// TIA Portal project "2023546359" (V18)

(* hardware
DEVICE "S7-1200 station_1"  S7-1200 Station
   slot 0: "Rack_0"  S7-1200 Rack  Rack  V1.0
   slot 1: "PLC"  CPU 1214C DC/DC/DC  6ES7 214-1AG40-0XB0  V4.2
*)

// ===== PLC "PLC"  CPU 1214C DC/DC/DC =====

VAR_GLOBAL CONSTANT   // PLC tag table "常量表"
   "ELE_SUM" : Int := 6;   // 电梯数量
   "FlOOR_TOP" : Int := 10;   // 电梯楼层
   "STATIC" : Int := 0;   // 静止状态
   "UP_H" : Int := 1;   // 上行高速
   "UP_L" : Int := 2;   // 上行低速
   "DOWN_H" : Int := 3;   // 下行高速
   "DOWN_L" : Int := 4;   // 下行低速
   "OPEN" : Int := 5;   // 开门
   "CLOSE" : Int := 6;   // 关门
   "H_L" : Int := 7;   // 高速转低速
   "L_H" : Int := 8;   // 低速转高速
   "SET_ELE" : Int := 5;
   "SET_FLOOR" : Int := 8;
END_VAR

TYPE "Button_Group"
   STRUCT
      state : Bool;
      light : Bool;
      p : Bool;
   END_STRUCT;
END_TYPE

TYPE "Elevator_Group"
   STRUCT
      jinggao : Struct
         REP : Bool;
         LC : Bool;
      END_STRUCT;
      display : Struct
         light : Bool;
         fan : Bool;
         error : Bool;
         full : Bool;
      END_STRUCT;
      direction : Struct
         up : Bool;
         down : Bool;
      END_STRUCT;
      door_jdq : Struct
         open : Bool;
         close : Bool;
      END_STRUCT;
      door_inplace : Struct
         close : Bool;
         open : Bool;
      END_STRUCT;
      bt_limit : Struct
         top1 : Bool;
         top2 : Bool;
         bottom1 : Bool;
         bottom2 : Bool;
      END_STRUCT;
      smg : Array[1..2, 1..7] of Bool;
      ele_speed : Struct
         H : Bool;
         L : Bool;
      END_STRUCT;
      run_contactor : Struct
         up : Bool;
         dowm : Bool;
      END_STRUCT;
      run_disp : Struct
         up : Bool;
         dowm : Bool;
      END_STRUCT;
      Brake : Struct
         B1 : Bool;
         B2 : Bool;
         B3 : Bool;
      END_STRUCT;
      floor_Lock : Array[1.."FlOOR_TOP"] of Bool;
      door_Lock : Bool;
      door_open : "Button_Group";
      btn_close : "Button_Group";
      ele_in_button : Array[1.."FlOOR_TOP"] of "Button_Group";
      run_enable : Bool;
      zhongliang : Word;
      button_out : Array[1..2, 1.."FlOOR_TOP"] of "Button_Group";   // 公共外部按键
   END_STRUCT;
END_TYPE

TYPE "Variable_Group"
   STRUCT
      init : Struct   // 初始化相关变量
         Init_state : Int;   // 初始化状态机
         kaishi : Bool;   // 初始化开始信号
         Init_now_f : Int;   // 初始化当前楼层
         mubiao_floor : Int;   // 初始化目标楼层
         init_fangxiang : Bool;   // 初始化方向
         jieshu : Bool;
         re_fangxiang : Bool;   // 检修后初始化方向
         re_mode : Bool;   // 检修后初始化方向设置模式(0自动1手动)
      END_STRUCT;
      Floor_handle : Struct   // 楼层处理相关变量
         dangqian_floor : Int;   // 当前楼层
         tag_1 : Bool;
         tag_2 : Bool;
      END_STRUCT;
      Weight_handle : Struct   // 重量处理相关变量
         m_load : Real;   // 标准化模拟量
         shiji_load : Real;   // 实际重量
         chaozhongxinhao : Bool;   // 超重信号
         jiangyao_chaozhong : Bool;   // 将要超载
         max_load : Real;   // 荷载重量
      END_STRUCT;
      yunxing_chuli : Struct   // 运行处理相关变量
         uopdown_state : Int;   // 上下行状态机
         run_state : Int;   // 运行状态机
         zuida_floor : Int;
         zuixiao_floor : Int;
         yunxu_run : Bool;   // 允许运行
      END_STRUCT;
      anniu_luru : Struct   // 内部按键录入变量
         neibu_anniu : Array[1.."FlOOR_TOP"] of Bool;
         waibu_anniu : Array[1..2, 0.."FlOOR_TOP"] of Bool;
      END_STRUCT;
      shijian : Array[1..13] of IEC_TIMER;   // 定时器变量
      Count : Array[1..3] of IEC_COUNTER;   // 计数器变量
      gaibian : Struct
         init_dir : Bool;   // 初始化方向
         init_aimf : Int;   // 初始化目标楼层
         max_load : Int;   // 荷载重量
         speed : Int;   // 电梯速度(1低2中3高)
         REP : Bool;   // 模拟检修信号
         now_load : Real;   // 模拟重量值
      END_STRUCT;
      qunkong : Struct   // 群控
         btn_time : Array[1.."FlOOR_TOP"] of Int;
         TH : Int;
      END_STRUCT;
      cuowu : Struct   // 异常处理
         stop : Bool;   // 特殊停层
         REP_deal : Bool;   // 检修处理
         tag_REPL : Bool;   // 检修处理下降沿检测
         tag_REPR : Bool;   // 检修处理上升沿检测
         start_cnt : Bool;   // 开始记录电梯异常状态
         error_time : Int;   // 处于异常状态时间
         qi_ting : Bool;
      END_STRUCT;
      interrupt : Struct
         state : Int;
         f_1ms : Bool;
         f_100ms : Bool;
         cnt_100ms : Int;
      END_STRUCT;
      报警指示灯 : Int;
      触发报警 : Int;
      状态指示灯 : Int;
      flag : Array[1..2, 0..10] of Bool;
   END_STRUCT;
END_TYPE

TYPE "Source"
   STRUCT
      MyBits : Struct
         btn_record : Array[1..32] of Bool;   // 总外呼按钮记录
         mainbtn_output : DWord;   // 总外呼输出
         state_record : Array[1..8] of Bool;   // 电梯状态记录
         state_output : Byte;   // 电梯状态输出
         floor_record : DWord;   // 楼层信号合并
         floor_record1 : Array[1..3] of DWord;   // 楼层信号输出
         btn_inside_record1 : Array[1..32] of Bool;   // 内呼按钮记录
         btn_inside_record2 : Array[1..32] of Bool;   // 内呼按钮记录
         btn_inside_record : Array[1..2] of DWord;   // 内呼按钮输出
         load_record : Array[1..3] of DWord;   // 载重记录输出
         start : Bool;   // 开始记录时间
         outsiedup1 : Array[1..32] of Bool;   // 虚拟外呼记录:1~3上呼
         outsiedup2 : Array[1..32] of Bool;   // 虚拟外呼记录:4~6上呼
         outsieddown1 : Array[1..32] of Bool;   // 虚拟外呼记录:1~3下呼
         outsieddown2 : Array[1..32] of Bool;   // 虚拟外呼记录:4~6下呼
         outside_fake : Array[1..4] of DWord;   // 虚拟外呼输出
         cnt_time : Int;   // 系统时间记录
      END_STRUCT;
   END_STRUCT;
END_TYPE

DATA_BLOCK "v_bianliang"   // DB1
{ S7_Optimized_Access := 'FALSE' }
VERSION : 0.1
   VAR
      dianti : Array[1.."ELE_SUM"] of "Variable_Group";
      anniu_waibu : Array[1..2, 0.."FlOOR_TOP"] of Bool;
      zidongyuxing_cnt : Int;   // 计算接受自动运行信号次数
      autorun : Bool;   // 模拟自动运行信号发生
      cnt_wancheng : Int;   // 计算完成初始化的电梯
      zuiyou_dianti : Int;   // 分配最优电梯
      mode_choice : Int;   // 模式选择
      time_min : Array[1.."ELE_SUM"] of Int;   // 候梯时间排序
      Source : "Source";
      interrupt : Struct
         f_1ms : Bool;
         cnt_100ms : Int;
         f_100ms : Bool;
      END_STRUCT;
      初始信号 : Bool;
      all_time : Struct
         sec : Int;
         min : Int;
         hour : Int;
         cnt_1s : Int;
      END_STRUCT;
      start_tim : Array[1..2, 1..10] of Int;
      over_tim : Array[1..2, 1..10] of Int;
      slope : Array[1..2, 1..10] of Real;
      zuiyou_louceng : Array[1..2] of Int;
      flag : Array[1..2] of Bool;
   END_VAR
BEGIN
   dianti[1].gaibian.speed := 3;
   dianti[1].gaibian.init_dir := 0;   // 初始化方向（0下1上）
   dianti[1].gaibian.init_aimf := 1;
   dianti[1].gaibian.max_load := 700;
   dianti[2].gaibian.init_aimf := 10;
   dianti[2].gaibian.max_load := 700;
   dianti[2].gaibian.speed := 3;
   dianti[3].gaibian.init_dir := 0;
   dianti[3].gaibian.init_aimf := 1;
   dianti[3].gaibian.max_load := 700;
   dianti[3].gaibian.speed := 3;
   time_min[1] := 0;
   time_min[2] := 0;
   time_min[3] := 0;
   dianti[2].gaibian.init_dir := 1;
   dianti[4].gaibian.init_dir := 0;
   dianti[4].gaibian.init_aimf := 1;
   dianti[4].gaibian.max_load := 700;
   dianti[4].gaibian.speed := 3;
   dianti[5].gaibian.init_dir := 0;
   dianti[5].gaibian.init_aimf := 1;
   dianti[5].gaibian.max_load := 1600;
   dianti[5].gaibian.speed := 2;
   dianti[6].gaibian.init_dir := 0;
   dianti[6].gaibian.init_aimf := 1;
   dianti[6].gaibian.max_load := 2000;
   dianti[6].gaibian.speed := 1;
   dianti[1].gaibian.REP := false;
   dianti[1].gaibian.now_load := 0.0;
   dianti[2].gaibian.REP := false;
   dianti[2].gaibian.now_load := 0.0;
   dianti[3].gaibian.REP := false;
   dianti[3].gaibian.now_load := 0.0;
   dianti[4].gaibian.REP := false;
   dianti[4].gaibian.now_load := 0.0;
   dianti[5].gaibian.REP := false;
   dianti[5].gaibian.now_load := 0.0;
   dianti[6].gaibian.REP := false;
   dianti[6].gaibian.now_load := 0.0;
   // dianti[1].anniu_luru.neibu_anniu : 响应按键
END_DATA_BLOCK

DATA_BLOCK "IO"   // DB2
{ S7_Optimized_Access := 'FALSE' }
VERSION : 0.1
   VAR
      software_autorun : Bool;   // 自动运行信号
      plc_ready : Bool;   // 准备就绪信号
      elev : Array[1.."ELE_SUM"] of "Elevator_Group";   // 电梯序号
   END_VAR
BEGIN
END_DATA_BLOCK

DATA_BLOCK "报警"   // DB5
{ S7_Optimized_Access := 'FALSE' }
VERSION : 0.1
   VAR
      维修报警 : Array[1..6] of Word;
      超重报警 : Array[1..6] of Word;
   END_VAR
BEGIN
END_DATA_BLOCK

DATA_BLOCK "INPUT"   // DB10
{ S7_Optimized_Access := 'FALSE' }
VERSION : 0.1
   VAR
      "1号梯1层上行呼梯按钮" : Bool;
      "1号梯2层上行呼梯按钮" : Bool;
      "1号梯3层上行呼梯按钮" : Bool;
      "1号梯4层上行呼梯按钮" : Bool;
      "1号梯5层上行呼梯按钮" : Bool;
      "1号梯6层上行呼梯按钮" : Bool;
      "1号梯7层上行呼梯按钮" : Bool;
      "1号梯8层上行呼梯按钮" : Bool;
      "1号梯9层上行呼梯按钮" : Bool;
      "1号梯2层下行呼梯按钮" : Bool;
      "1号梯3层下行呼梯按钮" : Bool;
      "1号梯4层下行呼梯按钮" : Bool;
      "1号梯5层下行呼梯按钮" : Bool;
      "1号梯6层下行呼梯按钮" : Bool;
      "1号梯7层下行呼梯按钮" : Bool;
      "1号梯8层下行呼梯按钮" : Bool;
      "1号梯9层下行呼梯按钮" : Bool;
      "1号梯10层下行呼梯按钮" : Bool;
      "1号梯轿内选层按钮1" : Bool;
      "1号梯轿内选层按钮2" : Bool;
      "1号梯轿内选层按钮3" : Bool;
      "1号梯轿内选层按钮4" : Bool;
      "1号梯轿内选层按钮5" : Bool;
      "1号梯轿内选层按钮6" : Bool;
      "1号梯轿内选层按钮7" : Bool;
      "1号梯轿内选层按钮8" : Bool;
      "1号梯轿内选层按钮9" : Bool;
      "1号梯轿内选层按钮10" : Bool;
      "1号梯轿内开门按钮" : Bool;
      "1号梯轿内关门按钮" : Bool;
      "1号梯光幕信号" : Bool;
      "1号梯检修信号" : Bool;
      "1号梯轿厢门锁信号" : Bool;
      "1号梯1楼层门锁信号" : Bool;
      "1号梯2楼层门锁信号" : Bool;
      "1号梯3楼层门锁信号" : Bool;
      "1号梯4楼层门锁信号" : Bool;
      "1号梯5楼层门锁信号" : Bool;
      "1号梯6楼层门锁信号" : Bool;
      "1号梯7楼层门锁信号" : Bool;
      "1号梯8楼层门锁信号" : Bool;
      "1号梯9楼层门锁信号" : Bool;
      "1号梯10楼层门锁信号" : Bool;
      "1号梯开门到位" : Bool;
      "1号梯关门到位" : Bool;
      "1号梯上平层信号" : Bool;
      "1号梯下平层信号" : Bool;
      "1号梯上端站第1限位" : Bool;
      "1号梯上端站第2限位" : Bool;
      "1号梯下端站第1限位" : Bool;
      "1号梯下端站第2限位" : Bool;
      "2号梯1层上行呼梯按钮" : Bool;
      "2号梯2层上行呼梯按钮" : Bool;
      "2号梯3层上行呼梯按钮" : Bool;
      "2号梯4层上行呼梯按钮" : Bool;
      "2号梯5层上行呼梯按钮" : Bool;
      "2号梯6层上行呼梯按钮" : Bool;
      "2号梯7层上行呼梯按钮" : Bool;
      "2号梯8层上行呼梯按钮" : Bool;
      "2号梯9层上行呼梯按钮" : Bool;
      "2号梯2层下行呼梯按钮" : Bool;
      "2号梯3层下行呼梯按钮" : Bool;
      "2号梯4层下行呼梯按钮" : Bool;
      "2号梯5层下行呼梯按钮" : Bool;
      "2号梯6层下行呼梯按钮" : Bool;
      "2号梯7层下行呼梯按钮" : Bool;
      "2号梯8层下行呼梯按钮" : Bool;
      "2号梯9层下行呼梯按钮" : Bool;
      "2号梯10层下行呼梯按钮" : Bool;
      "2号梯轿内选层按钮1" : Bool;
      "2号梯轿内选层按钮2" : Bool;
      "2号梯轿内选层按钮3" : Bool;
      "2号梯轿内选层按钮4" : Bool;
      "2号梯轿内选层按钮5" : Bool;
      "2号梯轿内选层按钮6" : Bool;
      "2号梯轿内选层按钮7" : Bool;
      "2号梯轿内选层按钮8" : Bool;
      "2号梯轿内选层按钮9" : Bool;
      "2号梯轿内选层按钮10" : Bool;
      "2号梯轿内开门按钮" : Bool;
      "2号梯轿内关门按钮" : Bool;
      "2号梯光幕信号" : Bool;
      "2号梯检修信号" : Bool;
      "2号梯轿厢门锁信号" : Bool;
      "2号梯1楼层门锁信号" : Bool;
      "2号梯2楼层门锁信号" : Bool;
      "2号梯3楼层门锁信号" : Bool;
      "2号梯4楼层门锁信号" : Bool;
      "2号梯5楼层门锁信号" : Bool;
      "2号梯6楼层门锁信号" : Bool;
      "2号梯7楼层门锁信号" : Bool;
      "2号梯8楼层门锁信号" : Bool;
      "2号梯9楼层门锁信号" : Bool;
      "2号梯10楼层门锁信号" : Bool;
      "2号梯开门到位" : Bool;
      "2号梯关门到位" : Bool;
      "2号梯上平层信号" : Bool;
      "2号梯下平层信号" : Bool;
      "2号梯上端站第1限位" : Bool;
      "2号梯上端站第2限位" : Bool;
      "2号梯下端站第1限位" : Bool;
      "2号梯下端站第2限位" : Bool;
      "3号梯1层上行呼梯按钮" : Bool;
      "3号梯2层上行呼梯按钮" : Bool;
      "3号梯3层上行呼梯按钮" : Bool;
      "3号梯4层上行呼梯按钮" : Bool;
      "3号梯5层上行呼梯按钮" : Bool;
      "3号梯6层上行呼梯按钮" : Bool;
      "3号梯7层上行呼梯按钮" : Bool;
      "3号梯8层上行呼梯按钮" : Bool;
      "3号梯9层上行呼梯按钮" : Bool;
      "3号梯2层下行呼梯按钮" : Bool;
      "3号梯3层下行呼梯按钮" : Bool;
      "3号梯4层下行呼梯按钮" : Bool;
      "3号梯5层下行呼梯按钮" : Bool;
      "3号梯6层下行呼梯按钮" : Bool;
      "3号梯7层下行呼梯按钮" : Bool;
      "3号梯8层下行呼梯按钮" : Bool;
      "3号梯9层下行呼梯按钮" : Bool;
      "3号梯10层下行呼梯按钮" : Bool;
      "3号梯轿内选层按钮1" : Bool;
      "3号梯轿内选层按钮2" : Bool;
      "3号梯轿内选层按钮3" : Bool;
      "3号梯轿内选层按钮4" : Bool;
      "3号梯轿内选层按钮5" : Bool;
      "3号梯轿内选层按钮6" : Bool;
      "3号梯轿内选层按钮7" : Bool;
      "3号梯轿内选层按钮8" : Bool;
      "3号梯轿内选层按钮9" : Bool;
      "3号梯轿内选层按钮10" : Bool;
      "3号梯轿内开门按钮" : Bool;
      "3号梯轿内关门按钮" : Bool;
      "3号梯光幕信号" : Bool;
      "3号梯检修信号" : Bool;
      "3号梯轿厢门锁信号" : Bool;
      "3号梯1楼层门锁信号" : Bool;
      "3号梯2楼层门锁信号" : Bool;
      "3号梯3楼层门锁信号" : Bool;
      "3号梯4楼层门锁信号" : Bool;
      "3号梯5楼层门锁信号" : Bool;
      "3号梯6楼层门锁信号" : Bool;
      "3号梯7楼层门锁信号" : Bool;
      "3号梯8楼层门锁信号" : Bool;
      "3号梯9楼层门锁信号" : Bool;
      "3号梯10楼层门锁信号" : Bool;
      "3号梯开门到位" : Bool;
      "3号梯关门到位" : Bool;
      "3号梯上平层信号" : Bool;
      "3号梯下平层信号" : Bool;
      "3号梯上端站第1限位" : Bool;
      "3号梯上端站第2限位" : Bool;
      "3号梯下端站第1限位" : Bool;
      "3号梯下端站第2限位" : Bool;
      "4号梯1层上行呼梯按钮" : Bool;
      "4号梯2层上行呼梯按钮" : Bool;
      "4号梯3层上行呼梯按钮" : Bool;
      "4号梯4层上行呼梯按钮" : Bool;
      "4号梯5层上行呼梯按钮" : Bool;
      "4号梯6层上行呼梯按钮" : Bool;
      "4号梯7层上行呼梯按钮" : Bool;
      "4号梯8层上行呼梯按钮" : Bool;
      "4号梯9层上行呼梯按钮" : Bool;
      "4号梯2层下行呼梯按钮" : Bool;
      "4号梯3层下行呼梯按钮" : Bool;
      "4号梯4层下行呼梯按钮" : Bool;
      "4号梯5层下行呼梯按钮" : Bool;
      "4号梯6层下行呼梯按钮" : Bool;
      "4号梯7层下行呼梯按钮" : Bool;
      "4号梯8层下行呼梯按钮" : Bool;
      "4号梯9层下行呼梯按钮" : Bool;
      "4号梯10层下行呼梯按钮" : Bool;
      "4号梯轿内选层按钮1" : Bool;
      "4号梯轿内选层按钮2" : Bool;
      "4号梯轿内选层按钮3" : Bool;
      "4号梯轿内选层按钮4" : Bool;
      "4号梯轿内选层按钮5" : Bool;
      "4号梯轿内选层按钮6" : Bool;
      "4号梯轿内选层按钮7" : Bool;
      "4号梯轿内选层按钮8" : Bool;
      "4号梯轿内选层按钮9" : Bool;
      "4号梯轿内选层按钮10" : Bool;
      "4号梯轿内开门按钮" : Bool;
      "4号梯轿内关门按钮" : Bool;
      "4号梯光幕信号" : Bool;
      "4号梯检修信号" : Bool;
      "4号梯轿厢门锁信号" : Bool;
      "4号梯1楼层门锁信号" : Bool;
      "4号梯2楼层门锁信号" : Bool;
      "4号梯3楼层门锁信号" : Bool;
      "4号梯4楼层门锁信号" : Bool;
      "4号梯5楼层门锁信号" : Bool;
      "4号梯6楼层门锁信号" : Bool;
      "4号梯7楼层门锁信号" : Bool;
      "4号梯8楼层门锁信号" : Bool;
      "4号梯9楼层门锁信号" : Bool;
      "4号梯10楼层门锁信号" : Bool;
      "4号梯开门到位" : Bool;
      "4号梯关门到位" : Bool;
      "4号梯上平层信号" : Bool;
      "4号梯下平层信号" : Bool;
      "4号梯上端站第1限位" : Bool;
      "4号梯上端站第2限位" : Bool;
      "4号梯下端站第1限位" : Bool;
      "4号梯下端站第2限位" : Bool;
      "5号梯1层上行呼梯按钮" : Bool;
      "5号梯2层上行呼梯按钮" : Bool;
      "5号梯3层上行呼梯按钮" : Bool;
      "5号梯4层上行呼梯按钮" : Bool;
      "5号梯5层上行呼梯按钮" : Bool;
      "5号梯6层上行呼梯按钮" : Bool;
      "5号梯7层上行呼梯按钮" : Bool;
      "5号梯8层上行呼梯按钮" : Bool;
      "5号梯9层上行呼梯按钮" : Bool;
      "5号梯2层下行呼梯按钮" : Bool;
      "5号梯3层下行呼梯按钮" : Bool;
      "5号梯4层下行呼梯按钮" : Bool;
      "5号梯5层下行呼梯按钮" : Bool;
      "5号梯6层下行呼梯按钮" : Bool;
      "5号梯7层下行呼梯按钮" : Bool;
      "5号梯8层下行呼梯按钮" : Bool;
      "5号梯9层下行呼梯按钮" : Bool;
      "5号梯10层下行呼梯按钮" : Bool;
      "5号梯轿内选层按钮1" : Bool;
      "5号梯轿内选层按钮2" : Bool;
      "5号梯轿内选层按钮3" : Bool;
      "5号梯轿内选层按钮4" : Bool;
      "5号梯轿内选层按钮5" : Bool;
      "5号梯轿内选层按钮6" : Bool;
      "5号梯轿内选层按钮7" : Bool;
      "5号梯轿内选层按钮8" : Bool;
      "5号梯轿内选层按钮9" : Bool;
      "5号梯轿内选层按钮10" : Bool;
      "5号梯轿内开门按钮" : Bool;
      "5号梯轿内关门按钮" : Bool;
      "5号梯光幕信号" : Bool;
      "5号梯检修信号" : Bool;
      "5号梯轿厢门锁信号" : Bool;
      "5号梯1楼层门锁信号" : Bool;
      "5号梯2楼层门锁信号" : Bool;
      "5号梯3楼层门锁信号" : Bool;
      "5号梯4楼层门锁信号" : Bool;
      "5号梯5楼层门锁信号" : Bool;
      "5号梯6楼层门锁信号" : Bool;
      "5号梯7楼层门锁信号" : Bool;
      "5号梯8楼层门锁信号" : Bool;
      "5号梯9楼层门锁信号" : Bool;
      "5号梯10楼层门锁信号" : Bool;
      "5号梯开门到位" : Bool;
      "5号梯关门到位" : Bool;
      "5号梯上平层信号" : Bool;
      "5号梯下平层信号" : Bool;
      "5号梯上端站第1限位" : Bool;
      "5号梯上端站第2限位" : Bool;
      "5号梯下端站第1限位" : Bool;
      "5号梯下端站第2限位" : Bool;
      "6号梯1层上行呼梯按钮" : Bool;
      "6号梯2层上行呼梯按钮" : Bool;
      "6号梯3层上行呼梯按钮" : Bool;
      "6号梯4层上行呼梯按钮" : Bool;
      "6号梯5层上行呼梯按钮" : Bool;
      "6号梯6层上行呼梯按钮" : Bool;
      "6号梯7层上行呼梯按钮" : Bool;
      "6号梯8层上行呼梯按钮" : Bool;
      "6号梯9层上行呼梯按钮" : Bool;
      "6号梯2层下行呼梯按钮" : Bool;
      "6号梯3层下行呼梯按钮" : Bool;
      "6号梯4层下行呼梯按钮" : Bool;
      "6号梯5层下行呼梯按钮" : Bool;
      "6号梯6层下行呼梯按钮" : Bool;
      "6号梯7层下行呼梯按钮" : Bool;
      "6号梯8层下行呼梯按钮" : Bool;
      "6号梯9层下行呼梯按钮" : Bool;
      "6号梯10层下行呼梯按钮" : Bool;
      "6号梯轿内选层按钮1" : Bool;
      "6号梯轿内选层按钮2" : Bool;
      "6号梯轿内选层按钮3" : Bool;
      "6号梯轿内选层按钮4" : Bool;
      "6号梯轿内选层按钮5" : Bool;
      "6号梯轿内选层按钮6" : Bool;
      "6号梯轿内选层按钮7" : Bool;
      "6号梯轿内选层按钮8" : Bool;
      "6号梯轿内选层按钮9" : Bool;
      "6号梯轿内选层按钮10" : Bool;
      "6号梯轿内开门按钮" : Bool;
      "6号梯轿内关门按钮" : Bool;
      "6号梯光幕信号" : Bool;
      "6号梯检修信号" : Bool;
      "6号梯轿厢门锁信号" : Bool;
      "6号梯1楼层门锁信号" : Bool;
      "6号梯2楼层门锁信号" : Bool;
      "6号梯3楼层门锁信号" : Bool;
      "6号梯4楼层门锁信号" : Bool;
      "6号梯5楼层门锁信号" : Bool;
      "6号梯6楼层门锁信号" : Bool;
      "6号梯7楼层门锁信号" : Bool;
      "6号梯8楼层门锁信号" : Bool;
      "6号梯9楼层门锁信号" : Bool;
      "6号梯10楼层门锁信号" : Bool;
      "6号梯开门到位" : Bool;
      "6号梯关门到位" : Bool;
      "6号梯上平层信号" : Bool;
      "6号梯下平层信号" : Bool;
      "6号梯上端站第1限位" : Bool;
      "6号梯上端站第2限位" : Bool;
      "6号梯下端站第1限位" : Bool;
      "6号梯下端站第2限位" : Bool;
      自动运行信号 : Bool;
      "1号梯当前载重量" : Word;
      "2号梯当前载重量" : Word;
      "3号梯当前载重量" : Word;
      "4号梯当前载重量" : Word;
      "5号梯当前载重量" : Word;
      "6号梯当前载重量" : Word;
   END_VAR
BEGIN
END_DATA_BLOCK

DATA_BLOCK "OUTPUT"   // DB11
{ S7_Optimized_Access := 'FALSE' }
VERSION : 0.1
   VAR
      "1号梯1层上行呼梯按钮指示灯" : Bool;
      "1号梯2层上行呼梯按钮指示灯" : Bool;
      "1号梯3层上行呼梯按钮指示灯" : Bool;
      "1号梯4层上行呼梯按钮指示灯" : Bool;
      "1号梯5层上行呼梯按钮指示灯" : Bool;
      "1号梯6层上行呼梯按钮指示灯" : Bool;
      "1号梯7层上行呼梯按钮指示灯" : Bool;
      "1号梯8层上行呼梯按钮指示灯" : Bool;
      "1号梯9层上行呼梯按钮指示灯" : Bool;
      "1号梯2层下行呼梯按钮指示灯" : Bool;
      "1号梯3层下行呼梯按钮指示灯" : Bool;
      "1号梯4层下行呼梯按钮指示灯" : Bool;
      "1号梯5层下行呼梯按钮指示灯" : Bool;
      "1号梯6层下行呼梯按钮指示灯" : Bool;
      "1号梯7层下行呼梯按钮指示灯" : Bool;
      "1号梯8层下行呼梯按钮指示灯" : Bool;
      "1号梯9层下行呼梯按钮指示灯" : Bool;
      "1号梯10层下行呼梯按钮指示灯" : Bool;
      "1号梯1层按钮指示灯" : Bool;
      "1号梯2层按钮指示灯" : Bool;
      "1号梯3层按钮指示灯" : Bool;
      "1号梯4层按钮指示灯" : Bool;
      "1号梯5层按钮指示灯" : Bool;
      "1号梯6层按钮指示灯" : Bool;
      "1号梯7层按钮指示灯" : Bool;
      "1号梯8层按钮指示灯" : Bool;
      "1号梯9层按钮指示灯" : Bool;
      "1号梯10层按钮指示灯" : Bool;
      "1号梯LEDa" : Bool;
      "1号梯LEDb" : Bool;
      "1号梯LEDc" : Bool;
      "1号梯LEDd" : Bool;
      "1号梯LEDe" : Bool;
      "1号梯LEDf" : Bool;
      "1号梯LEDg" : Bool;
      "1号梯LEDh" : Bool;
      "1号梯LEDi" : Bool;
      "1号梯LEDj" : Bool;
      "1号梯LEDk" : Bool;
      "1号梯LEDl" : Bool;
      "1号梯LEDm" : Bool;
      "1号梯LEDn" : Bool;
      "1号梯上行指示" : Bool;
      "1号梯下行指示" : Bool;
      "1号梯故障指示" : Bool;
      "1号梯照明指示" : Bool;
      "1号梯风扇指示" : Bool;
      "1号梯满载指示" : Bool;
      "1号梯电机启动信号" : Bool;
      "1号梯上行接触器" : Bool;
      "1号梯下行接触器" : Bool;
      "1号梯高速接触器" : Bool;
      "1号梯低速接触器" : Bool;
      "1号梯开门继电器" : Bool;
      "1号梯关门继电器" : Bool;
      "1号梯1级减速制动" : Bool;
      "1号梯2级减速制动" : Bool;
      "1号梯3级减速制动" : Bool;
      "2号梯1层上行呼梯按钮指示灯" : Bool;
      "2号梯2层上行呼梯按钮指示灯" : Bool;
      "2号梯3层上行呼梯按钮指示灯" : Bool;
      "2号梯4层上行呼梯按钮指示灯" : Bool;
      "2号梯5层上行呼梯按钮指示灯" : Bool;
      "2号梯6层上行呼梯按钮指示灯" : Bool;
      "2号梯7层上行呼梯按钮指示灯" : Bool;
      "2号梯8层上行呼梯按钮指示灯" : Bool;
      "2号梯9层上行呼梯按钮指示灯" : Bool;
      "2号梯2层下行呼梯按钮指示灯" : Bool;
      "2号梯3层下行呼梯按钮指示灯" : Bool;
      "2号梯4层下行呼梯按钮指示灯" : Bool;
      "2号梯5层下行呼梯按钮指示灯" : Bool;
      "2号梯6层下行呼梯按钮指示灯" : Bool;
      "2号梯7层下行呼梯按钮指示灯" : Bool;
      "2号梯8层下行呼梯按钮指示灯" : Bool;
      "2号梯9层下行呼梯按钮指示灯" : Bool;
      "2号梯10层下行呼梯按钮指示灯" : Bool;
      "2号梯1层按钮指示灯" : Bool;
      "2号梯2层按钮指示灯" : Bool;
      "2号梯3层按钮指示灯" : Bool;
      "2号梯4层按钮指示灯" : Bool;
      "2号梯5层按钮指示灯" : Bool;
      "2号梯6层按钮指示灯" : Bool;
      "2号梯7层按钮指示灯" : Bool;
      "2号梯8层按钮指示灯" : Bool;
      "2号梯9层按钮指示灯" : Bool;
      "2号梯10层按钮指示灯" : Bool;
      "2号梯LEDa" : Bool;
      "2号梯LEDb" : Bool;
      "2号梯LEDc" : Bool;
      "2号梯LEDd" : Bool;
      "2号梯LEDe" : Bool;
      "2号梯LEDf" : Bool;
      "2号梯LEDg" : Bool;
      "2号梯LEDh" : Bool;
      "2号梯LEDi" : Bool;
      "2号梯LEDj" : Bool;
      "2号梯LEDk" : Bool;
      "2号梯LEDl" : Bool;
      "2号梯LEDm" : Bool;
      "2号梯LEDn" : Bool;
      "2号梯上行指示" : Bool;
      "2号梯下行指示" : Bool;
      "2号梯故障指示" : Bool;
      "2号梯照明指示" : Bool;
      "2号梯风扇指示" : Bool;
      "2号梯满载指示" : Bool;
      "2号梯电机启动信号" : Bool;
      "2号梯上行接触器" : Bool;
      "2号梯下行接触器" : Bool;
      "2号梯高速接触器" : Bool;
      "2号梯低速接触器" : Bool;
      "2号梯开门继电器" : Bool;
      "2号梯关门继电器" : Bool;
      "2号梯1级减速制动" : Bool;
      "2号梯2级减速制动" : Bool;
      "2号梯3级减速制动" : Bool;
      "3号梯1层上行呼梯按钮指示灯" : Bool;
      "3号梯2层上行呼梯按钮指示灯" : Bool;
      "3号梯3层上行呼梯按钮指示灯" : Bool;
      "3号梯4层上行呼梯按钮指示灯" : Bool;
      "3号梯5层上行呼梯按钮指示灯" : Bool;
      "3号梯6层上行呼梯按钮指示灯" : Bool;
      "3号梯7层上行呼梯按钮指示灯" : Bool;
      "3号梯8层上行呼梯按钮指示灯" : Bool;
      "3号梯9层上行呼梯按钮指示灯" : Bool;
      "3号梯2层下行呼梯按钮指示灯" : Bool;
      "3号梯3层下行呼梯按钮指示灯" : Bool;
      "3号梯4层下行呼梯按钮指示灯" : Bool;
      "3号梯5层下行呼梯按钮指示灯" : Bool;
      "3号梯6层下行呼梯按钮指示灯" : Bool;
      "3号梯7层下行呼梯按钮指示灯" : Bool;
      "3号梯8层下行呼梯按钮指示灯" : Bool;
      "3号梯9层下行呼梯按钮指示灯" : Bool;
      "3号梯10层下行呼梯按钮指示灯" : Bool;
      "3号梯1层按钮指示灯" : Bool;
      "3号梯2层按钮指示灯" : Bool;
      "3号梯3层按钮指示灯" : Bool;
      "3号梯4层按钮指示灯" : Bool;
      "3号梯5层按钮指示灯" : Bool;
      "3号梯6层按钮指示灯" : Bool;
      "3号梯7层按钮指示灯" : Bool;
      "3号梯8层按钮指示灯" : Bool;
      "3号梯9层按钮指示灯" : Bool;
      "3号梯10层按钮指示灯" : Bool;
      "3号梯LEDa" : Bool;
      "3号梯LEDb" : Bool;
      "3号梯LEDc" : Bool;
      "3号梯LEDd" : Bool;
      "3号梯LEDe" : Bool;
      "3号梯LEDf" : Bool;
      "3号梯LEDg" : Bool;
      "3号梯LEDh" : Bool;
      "3号梯LEDi" : Bool;
      "3号梯LEDj" : Bool;
      "3号梯LEDk" : Bool;
      "3号梯LEDl" : Bool;
      "3号梯LEDm" : Bool;
      "3号梯LEDn" : Bool;
      "3号梯上行指示" : Bool;
      "3号梯下行指示" : Bool;
      "3号梯故障指示" : Bool;
      "3号梯照明指示" : Bool;
      "3号梯风扇指示" : Bool;
      "3号梯满载指示" : Bool;
      "3号梯电机启动信号" : Bool;
      "3号梯上行接触器" : Bool;
      "3号梯下行接触器" : Bool;
      "3号梯高速接触器" : Bool;
      "3号梯低速接触器" : Bool;
      "3号梯开门继电器" : Bool;
      "3号梯关门继电器" : Bool;
      "3号梯1级减速制动" : Bool;
      "3号梯2级减速制动" : Bool;
      "3号梯3级减速制动" : Bool;
      "4号梯1层上行呼梯按钮指示灯" : Bool;
      "4号梯2层上行呼梯按钮指示灯" : Bool;
      "4号梯3层上行呼梯按钮指示灯" : Bool;
      "4号梯4层上行呼梯按钮指示灯" : Bool;
      "4号梯5层上行呼梯按钮指示灯" : Bool;
      "4号梯6层上行呼梯按钮指示灯" : Bool;
      "4号梯7层上行呼梯按钮指示灯" : Bool;
      "4号梯8层上行呼梯按钮指示灯" : Bool;
      "4号梯9层上行呼梯按钮指示灯" : Bool;
      "4号梯2层下行呼梯按钮指示灯" : Bool;
      "4号梯3层下行呼梯按钮指示灯" : Bool;
      "4号梯4层下行呼梯按钮指示灯" : Bool;
      "4号梯5层下行呼梯按钮指示灯" : Bool;
      "4号梯6层下行呼梯按钮指示灯" : Bool;
      "4号梯7层下行呼梯按钮指示灯" : Bool;
      "4号梯8层下行呼梯按钮指示灯" : Bool;
      "4号梯9层下行呼梯按钮指示灯" : Bool;
      "4号梯10层下行呼梯按钮指示灯" : Bool;
      "4号梯1层按钮指示灯" : Bool;
      "4号梯2层按钮指示灯" : Bool;
      "4号梯3层按钮指示灯" : Bool;
      "4号梯4层按钮指示灯" : Bool;
      "4号梯5层按钮指示灯" : Bool;
      "4号梯6层按钮指示灯" : Bool;
      "4号梯7层按钮指示灯" : Bool;
      "4号梯8层按钮指示灯" : Bool;
      "4号梯9层按钮指示灯" : Bool;
      "4号梯10层按钮指示灯" : Bool;
      "4号梯LEDa" : Bool;
      "4号梯LEDb" : Bool;
      "4号梯LEDc" : Bool;
      "4号梯LEDd" : Bool;
      "4号梯LEDe" : Bool;
      "4号梯LEDf" : Bool;
      "4号梯LEDg" : Bool;
      "4号梯LEDh" : Bool;
      "4号梯LEDi" : Bool;
      "4号梯LEDj" : Bool;
      "4号梯LEDk" : Bool;
      "4号梯LEDl" : Bool;
      "4号梯LEDm" : Bool;
      "4号梯LEDn" : Bool;
      "4号梯上行指示" : Bool;
      "4号梯下行指示" : Bool;
      "4号梯故障指示" : Bool;
      "4号梯照明指示" : Bool;
      "4号梯风扇指示" : Bool;
      "4号梯满载指示" : Bool;
      "4号梯电机启动信号" : Bool;
      "4号梯上行接触器" : Bool;
      "4号梯下行接触器" : Bool;
      "4号梯高速接触器" : Bool;
      "4号梯低速接触器" : Bool;
      "4号梯开门继电器" : Bool;
      "4号梯关门继电器" : Bool;
      "4号梯1级减速制动" : Bool;
      "4号梯2级减速制动" : Bool;
      "4号梯3级减速制动" : Bool;
      "5号梯1层上行呼梯按钮指示灯" : Bool;
      "5号梯2层上行呼梯按钮指示灯" : Bool;
      "5号梯3层上行呼梯按钮指示灯" : Bool;
      "5号梯4层上行呼梯按钮指示灯" : Bool;
      "5号梯5层上行呼梯按钮指示灯" : Bool;
      "5号梯6层上行呼梯按钮指示灯" : Bool;
      "5号梯7层上行呼梯按钮指示灯" : Bool;
      "5号梯8层上行呼梯按钮指示灯" : Bool;
      "5号梯9层上行呼梯按钮指示灯" : Bool;
      "5号梯2层下行呼梯按钮指示灯" : Bool;
      "5号梯3层下行呼梯按钮指示灯" : Bool;
      "5号梯4层下行呼梯按钮指示灯" : Bool;
      "5号梯5层下行呼梯按钮指示灯" : Bool;
      "5号梯6层下行呼梯按钮指示灯" : Bool;
      "5号梯7层下行呼梯按钮指示灯" : Bool;
      "5号梯8层下行呼梯按钮指示灯" : Bool;
      "5号梯9层下行呼梯按钮指示灯" : Bool;
      "5号梯10层下行呼梯按钮指示灯" : Bool;
      "5号梯1层按钮指示灯" : Bool;
      "5号梯2层按钮指示灯" : Bool;
      "5号梯3层按钮指示灯" : Bool;
      "5号梯4层按钮指示灯" : Bool;
      "5号梯5层按钮指示灯" : Bool;
      "5号梯6层按钮指示灯" : Bool;
      "5号梯7层按钮指示灯" : Bool;
      "5号梯8层按钮指示灯" : Bool;
      "5号梯9层按钮指示灯" : Bool;
      "5号梯10层按钮指示灯" : Bool;
      "5号梯LEDa" : Bool;
      "5号梯LEDb" : Bool;
      "5号梯LEDc" : Bool;
      "5号梯LEDd" : Bool;
      "5号梯LEDe" : Bool;
      "5号梯LEDf" : Bool;
      "5号梯LEDg" : Bool;
      "5号梯LEDh" : Bool;
      "5号梯LEDi" : Bool;
      "5号梯LEDj" : Bool;
      "5号梯LEDk" : Bool;
      "5号梯LEDl" : Bool;
      "5号梯LEDm" : Bool;
      "5号梯LEDn" : Bool;
      "5号梯上行指示" : Bool;
      "5号梯下行指示" : Bool;
      "5号梯故障指示" : Bool;
      "5号梯照明指示" : Bool;
      "5号梯风扇指示" : Bool;
      "5号梯满载指示" : Bool;
      "5号梯电机启动信号" : Bool;
      "5号梯上行接触器" : Bool;
      "5号梯下行接触器" : Bool;
      "5号梯高速接触器" : Bool;
      "5号梯低速接触器" : Bool;
      "5号梯开门继电器" : Bool;
      "5号梯关门继电器" : Bool;
      "5号梯1级减速制动" : Bool;
      "5号梯2级减速制动" : Bool;
      "5号梯3级减速制动" : Bool;
      "6号梯1层上行呼梯按钮指示灯" : Bool;
      "6号梯2层上行呼梯按钮指示灯" : Bool;
      "6号梯3层上行呼梯按钮指示灯" : Bool;
      "6号梯4层上行呼梯按钮指示灯" : Bool;
      "6号梯5层上行呼梯按钮指示灯" : Bool;
      "6号梯6层上行呼梯按钮指示灯" : Bool;
      "6号梯7层上行呼梯按钮指示灯" : Bool;
      "6号梯8层上行呼梯按钮指示灯" : Bool;
      "6号梯9层上行呼梯按钮指示灯" : Bool;
      "6号梯2层下行呼梯按钮指示灯" : Bool;
      "6号梯3层下行呼梯按钮指示灯" : Bool;
      "6号梯4层下行呼梯按钮指示灯" : Bool;
      "6号梯5层下行呼梯按钮指示灯" : Bool;
      "6号梯6层下行呼梯按钮指示灯" : Bool;
      "6号梯7层下行呼梯按钮指示灯" : Bool;
      "6号梯8层下行呼梯按钮指示灯" : Bool;
      "6号梯9层下行呼梯按钮指示灯" : Bool;
      "6号梯10层下行呼梯按钮指示灯" : Bool;
      "6号梯1层按钮指示灯" : Bool;
      "6号梯2层按钮指示灯" : Bool;
      "6号梯3层按钮指示灯" : Bool;
      "6号梯4层按钮指示灯" : Bool;
      "6号梯5层按钮指示灯" : Bool;
      "6号梯6层按钮指示灯" : Bool;
      "6号梯7层按钮指示灯" : Bool;
      "6号梯8层按钮指示灯" : Bool;
      "6号梯9层按钮指示灯" : Bool;
      "6号梯10层按钮指示灯" : Bool;
      "6号梯LEDa" : Bool;
      "6号梯LEDb" : Bool;
      "6号梯LEDc" : Bool;
      "6号梯LEDd" : Bool;
      "6号梯LEDe" : Bool;
      "6号梯LEDf" : Bool;
      "6号梯LEDg" : Bool;
      "6号梯LEDh" : Bool;
      "6号梯LEDi" : Bool;
      "6号梯LEDj" : Bool;
      "6号梯LEDk" : Bool;
      "6号梯LEDl" : Bool;
      "6号梯LEDm" : Bool;
      "6号梯LEDn" : Bool;
      "6号梯上行指示" : Bool;
      "6号梯下行指示" : Bool;
      "6号梯故障指示" : Bool;
      "6号梯照明指示" : Bool;
      "6号梯风扇指示" : Bool;
      "6号梯满载指示" : Bool;
      "6号梯电机启动信号" : Bool;
      "6号梯上行接触器" : Bool;
      "6号梯下行接触器" : Bool;
      "6号梯高速接触器" : Bool;
      "6号梯低速接触器" : Bool;
      "6号梯开门继电器" : Bool;
      "6号梯关门继电器" : Bool;
      "6号梯1级减速制动" : Bool;
      "6号梯2级减速制动" : Bool;
      "6号梯3级减速制动" : Bool;
      准备就绪信号 : Bool;
   END_VAR
BEGIN
END_DATA_BLOCK

FUNCTION "addr management" : Void   // FC1, SCL
{ S7_Optimized_Access := 'TRUE' }
VERSION : 0.1
BEGIN
   //地址映射
   //************************************************************************************************************************//
   //***********************************************INPUT********************************************************************//
   REGION 公共部分
       "IO".software_autorun := "INPUT".自动运行信号;

   END_REGION
   REGION 1号梯INPUT 
       "IO".elev[1].ele_in_button[1].state := "INPUT"."1号梯轿内选层按钮1";
       "IO".elev[1].ele_in_button[2].state := "INPUT"."1号梯轿内选层按钮2";
       "IO".elev[1].ele_in_button[3].state := "INPUT"."1号梯轿内选层按钮3";
       "IO".elev[1].ele_in_button[4].state := "INPUT"."1号梯轿内选层按钮4";
       "IO".elev[1].ele_in_button[5].state := "INPUT"."1号梯轿内选层按钮5";
       "IO".elev[1].ele_in_button[6].state := "INPUT"."1号梯轿内选层按钮6";
       "IO".elev[1].ele_in_button[7].state := "INPUT"."1号梯轿内选层按钮7";
       "IO".elev[1].ele_in_button[8].state := "INPUT"."1号梯轿内选层按钮8";
       "IO".elev[1].ele_in_button[9].state := "INPUT"."1号梯轿内选层按钮9";
       "IO".elev[1].ele_in_button[10].state := "INPUT"."1号梯轿内选层按钮10";

       "IO".elev[1].door_open.state := "INPUT"."1号梯轿内开门按钮";
       "IO".elev[1].btn_close.state := "INPUT"."1号梯轿内关门按钮";

       "IO".elev[1].door_Lock := "INPUT"."1号梯轿厢门锁信号";
       "IO".elev[1].floor_Lock[1] := "INPUT"."1号梯1楼层门锁信号";
       "IO".elev[1].floor_Lock[2] := "INPUT"."1号梯2楼层门锁信号";
       "IO".elev[1].floor_Lock[3] := "INPUT"."1号梯3楼层门锁信号";
       "IO".elev[1].floor_Lock[4] := "INPUT"."1号梯4楼层门锁信号";
       "IO".elev[1].floor_Lock[5] := "INPUT"."1号梯5楼层门锁信号";
       "IO".elev[1].floor_Lock[6] := "INPUT"."1号梯6楼层门锁信号";
       "IO".elev[1].floor_Lock[7] := "INPUT"."1号梯7楼层门锁信号";
       "IO".elev[1].floor_Lock[8] := "INPUT"."1号梯8楼层门锁信号";
       "IO".elev[1].floor_Lock[9] := "INPUT"."1号梯9楼层门锁信号";
       "IO".elev[1].floor_Lock[10] := "INPUT"."1号梯10楼层门锁信号";

       "IO".elev[1].button_out[1, 1].state := "INPUT"."1号梯1层上行呼梯按钮";
       "IO".elev[1].button_out[1, 2].state := "INPUT"."1号梯2层上行呼梯按钮";
       "IO".elev[1].button_out[1, 3].state := "INPUT"."1号梯3层上行呼梯按钮";
       "IO".elev[1].button_out[1, 4].state := "INPUT"."1号梯4层上行呼梯按钮";
       "IO".elev[1].button_out[1, 5].state := "INPUT"."1号梯5层上行呼梯按钮";
       "IO".elev[1].button_out[1, 6].state := "INPUT"."1号梯6层上行呼梯按钮";
       "IO".elev[1].button_out[1, 7].state := "INPUT"."1号梯7层上行呼梯按钮";
       "IO".elev[1].button_out[1, 8].state := "INPUT"."1号梯8层上行呼梯按钮";
       "IO".elev[1].button_out[1, 9].state := "INPUT"."1号梯9层上行呼梯按钮";

       "IO".elev[1].button_out[2, 2].state := "INPUT"."1号梯2层下行呼梯按钮";
       "IO".elev[1].button_out[2, 3].state := "INPUT"."1号梯3层下行呼梯按钮";
       "IO".elev[1].button_out[2, 4].state := "INPUT"."1号梯4层下行呼梯按钮";
       "IO".elev[1].button_out[2, 5].state := "INPUT"."1号梯5层下行呼梯按钮";
       "IO".elev[1].button_out[2, 6].state := "INPUT"."1号梯6层下行呼梯按钮";
       "IO".elev[1].button_out[2, 7].state := "INPUT"."1号梯7层下行呼梯按钮";
       "IO".elev[1].button_out[2, 8].state := "INPUT"."1号梯8层下行呼梯按钮";
       "IO".elev[1].button_out[2, 9].state := "INPUT"."1号梯9层下行呼梯按钮";
       "IO".elev[1].button_out[2, 10].state := "INPUT"."1号梯10层下行呼梯按钮";

       "IO".elev[1].door_inplace.open := "INPUT"."1号梯开门到位";
       "IO".elev[1].door_inplace.close := "INPUT"."1号梯关门到位";

       "IO".elev[1].direction.up := "INPUT"."1号梯上平层信号";
       "IO".elev[1].direction.down := "INPUT"."1号梯下平层信号";

       "IO".elev[1].jinggao.LC := "INPUT"."1号梯光幕信号";
       "IO".elev[1].jinggao.REP := "INPUT"."1号梯检修信号";

       "IO".elev[1].bt_limit.bottom1 := "INPUT"."1号梯下端站第1限位";
       "IO".elev[1].bt_limit.bottom2 := "INPUT"."1号梯下端站第2限位";
       "IO".elev[1].bt_limit.top1 := "INPUT"."1号梯上端站第1限位";
       "IO".elev[1].bt_limit.top2 := "INPUT"."1号梯上端站第2限位";

       "IO".elev[1].zhongliang := "INPUT"."1号梯当前载重量";
   END_REGION
   REGION 2号梯INPUT
       "IO".elev[2].ele_in_button[1].state := "INPUT"."2号梯轿内选层按钮1";
       "IO".elev[2].ele_in_button[2].state := "INPUT"."2号梯轿内选层按钮2";
       "IO".elev[2].ele_in_button[3].state := "INPUT"."2号梯轿内选层按钮3";
       "IO".elev[2].ele_in_button[4].state := "INPUT"."2号梯轿内选层按钮4";
       "IO".elev[2].ele_in_button[5].state := "INPUT"."2号梯轿内选层按钮5";
       "IO".elev[2].ele_in_button[6].state := "INPUT"."2号梯轿内选层按钮6";
       "IO".elev[2].ele_in_button[7].state := "INPUT"."2号梯轿内选层按钮7";
       "IO".elev[2].ele_in_button[8].state := "INPUT"."2号梯轿内选层按钮8";
       "IO".elev[2].ele_in_button[9].state := "INPUT"."2号梯轿内选层按钮9";
       "IO".elev[2].ele_in_button[10].state := "INPUT"."2号梯轿内选层按钮10";

       "IO".elev[2].door_open.state := "INPUT"."2号梯轿内开门按钮";
       "IO".elev[2].btn_close.state := "INPUT"."2号梯轿内关门按钮";

       "IO".elev[2].door_Lock := "INPUT"."2号梯轿厢门锁信号";
       "IO".elev[2].floor_Lock[1] := "INPUT"."2号梯1楼层门锁信号";
       "IO".elev[2].floor_Lock[2] := "INPUT"."2号梯2楼层门锁信号";
       "IO".elev[2].floor_Lock[3] := "INPUT"."2号梯3楼层门锁信号";
       "IO".elev[2].floor_Lock[4] := "INPUT"."2号梯4楼层门锁信号";
       "IO".elev[2].floor_Lock[5] := "INPUT"."2号梯5楼层门锁信号";
       "IO".elev[2].floor_Lock[6] := "INPUT"."2号梯6楼层门锁信号";
       "IO".elev[2].floor_Lock[7] := "INPUT"."2号梯7楼层门锁信号";
       "IO".elev[2].floor_Lock[8] := "INPUT"."2号梯8楼层门锁信号";
       "IO".elev[2].floor_Lock[9] := "INPUT"."2号梯9楼层门锁信号";
       "IO".elev[2].floor_Lock[10] := "INPUT"."2号梯10楼层门锁信号";

       "IO".elev[2].button_out[1, 1].state := "INPUT"."2号梯1层上行呼梯按钮";
       "IO".elev[2].button_out[1, 2].state := "INPUT"."2号梯2层上行呼梯按钮";
       "IO".elev[2].button_out[1, 3].state := "INPUT"."2号梯3层上行呼梯按钮";
       "IO".elev[2].button_out[1, 4].state := "INPUT"."2号梯4层上行呼梯按钮";
       "IO".elev[2].button_out[1, 5].state := "INPUT"."2号梯5层上行呼梯按钮";
       "IO".elev[2].button_out[1, 6].state := "INPUT"."2号梯6层上行呼梯按钮";
       "IO".elev[2].button_out[1, 7].state := "INPUT"."2号梯7层上行呼梯按钮";
       "IO".elev[2].button_out[1, 8].state := "INPUT"."2号梯8层上行呼梯按钮";
       "IO".elev[2].button_out[1, 9].state := "INPUT"."2号梯9层上行呼梯按钮";

       "IO".elev[2].button_out[2, 2].state := "INPUT"."2号梯2层下行呼梯按钮";
       "IO".elev[2].button_out[2, 3].state := "INPUT"."2号梯3层下行呼梯按钮";
       "IO".elev[2].button_out[2, 4].state := "INPUT"."2号梯4层下行呼梯按钮";
       "IO".elev[2].button_out[2, 5].state := "INPUT"."2号梯5层下行呼梯按钮";
       "IO".elev[2].button_out[2, 6].state := "INPUT"."2号梯6层下行呼梯按钮";
       "IO".elev[2].button_out[2, 7].state := "INPUT"."2号梯7层下行呼梯按钮";
       "IO".elev[2].button_out[2, 8].state := "INPUT"."2号梯8层下行呼梯按钮";
       "IO".elev[2].button_out[2, 9].state := "INPUT"."2号梯9层下行呼梯按钮";
       "IO".elev[2].button_out[2, 10].state := "INPUT"."2号梯10层下行呼梯按钮";

       "IO".elev[2].door_inplace.open := "INPUT"."2号梯开门到位";
       "IO".elev[2].door_inplace.close := "INPUT"."2号梯关门到位";

       "IO".elev[2].direction.up := "INPUT"."2号梯上平层信号";
       "IO".elev[2].direction.down := "INPUT"."2号梯下平层信号";

       "IO".elev[2].jinggao.LC := "INPUT"."2号梯光幕信号";
       "IO".elev[2].jinggao.REP := "INPUT"."2号梯检修信号";

       "IO".elev[2].bt_limit.bottom1 := "INPUT"."2号梯下端站第1限位";
       "IO".elev[2].bt_limit.bottom2 := "INPUT"."2号梯下端站第2限位";
       "IO".elev[2].bt_limit.top1 := "INPUT"."2号梯上端站第1限位";
       "IO".elev[2].bt_limit.top2 := "INPUT"."2号梯上端站第2限位";

       "IO".elev[2].zhongliang := "INPUT"."2号梯当前载重量";
   END_REGION
   REGION 3号梯INPUT
       "IO".elev[3].ele_in_button[1].state := "INPUT"."3号梯轿内选层按钮1";
       "IO".elev[3].ele_in_button[2].state := "INPUT"."3号梯轿内选层按钮2";
       "IO".elev[3].ele_in_button[3].state := "INPUT"."3号梯轿内选层按钮3";
       "IO".elev[3].ele_in_button[4].state := "INPUT"."3号梯轿内选层按钮4";
       "IO".elev[3].ele_in_button[5].state := "INPUT"."3号梯轿内选层按钮5";
       "IO".elev[3].ele_in_button[6].state := "INPUT"."3号梯轿内选层按钮6";
       "IO".elev[3].ele_in_button[7].state := "INPUT"."3号梯轿内选层按钮7";
       "IO".elev[3].ele_in_button[8].state := "INPUT"."3号梯轿内选层按钮8";
       "IO".elev[3].ele_in_button[9].state := "INPUT"."3号梯轿内选层按钮9";
       "IO".elev[3].ele_in_button[10].state := "INPUT"."3号梯轿内选层按钮10";

       "IO".elev[3].door_open.state := "INPUT"."3号梯轿内开门按钮";
       "IO".elev[3].btn_close.state := "INPUT"."3号梯轿内关门按钮";

       "IO".elev[3].door_Lock := "INPUT"."3号梯轿厢门锁信号";
       "IO".elev[3].floor_Lock[1] := "INPUT"."3号梯1楼层门锁信号";
       "IO".elev[3].floor_Lock[2] := "INPUT"."3号梯2楼层门锁信号";
       "IO".elev[3].floor_Lock[3] := "INPUT"."3号梯3楼层门锁信号";
       "IO".elev[3].floor_Lock[4] := "INPUT"."3号梯4楼层门锁信号";
       "IO".elev[3].floor_Lock[5] := "INPUT"."3号梯5楼层门锁信号";
       "IO".elev[3].floor_Lock[6] := "INPUT"."3号梯6楼层门锁信号";
       "IO".elev[3].floor_Lock[7] := "INPUT"."3号梯7楼层门锁信号";
       "IO".elev[3].floor_Lock[8] := "INPUT"."3号梯8楼层门锁信号";
       "IO".elev[3].floor_Lock[9] := "INPUT"."3号梯9楼层门锁信号";
       "IO".elev[3].floor_Lock[10] := "INPUT"."3号梯10楼层门锁信号";

       "IO".elev[3].button_out[1, 1].state := "INPUT"."3号梯1层上行呼梯按钮";
       "IO".elev[3].button_out[1, 2].state := "INPUT"."3号梯2层上行呼梯按钮";
       "IO".elev[3].button_out[1, 3].state := "INPUT"."3号梯3层上行呼梯按钮";
       "IO".elev[3].button_out[1, 4].state := "INPUT"."3号梯4层上行呼梯按钮";
       "IO".elev[3].button_out[1, 5].state := "INPUT"."3号梯5层上行呼梯按钮";
       "IO".elev[3].button_out[1, 6].state := "INPUT"."3号梯6层上行呼梯按钮";
       "IO".elev[3].button_out[1, 7].state := "INPUT"."3号梯7层上行呼梯按钮";
       "IO".elev[3].button_out[1, 8].state := "INPUT"."3号梯8层上行呼梯按钮";
       "IO".elev[3].button_out[1, 9].state := "INPUT"."3号梯9层上行呼梯按钮";

       "IO".elev[3].button_out[2, 2].state := "INPUT"."3号梯2层下行呼梯按钮";
       "IO".elev[3].button_out[2, 3].state := "INPUT"."3号梯3层下行呼梯按钮";
       "IO".elev[3].button_out[2, 4].state := "INPUT"."3号梯4层下行呼梯按钮";
       "IO".elev[3].button_out[2, 5].state := "INPUT"."3号梯5层下行呼梯按钮";
       "IO".elev[3].button_out[2, 6].state := "INPUT"."3号梯6层下行呼梯按钮";
       "IO".elev[3].button_out[2, 7].state := "INPUT"."3号梯7层下行呼梯按钮";
       "IO".elev[3].button_out[2, 8].state := "INPUT"."3号梯8层下行呼梯按钮";
       "IO".elev[3].button_out[2, 9].state := "INPUT"."3号梯9层下行呼梯按钮";
       "IO".elev[3].button_out[2, 10].state := "INPUT"."3号梯10层下行呼梯按钮";

       "IO".elev[3].door_inplace.open := "INPUT"."3号梯开门到位";
       "IO".elev[3].door_inplace.close := "INPUT"."3号梯关门到位";

       "IO".elev[3].direction.up := "INPUT"."3号梯上平层信号";
       "IO".elev[3].direction.down := "INPUT"."3号梯下平层信号";

       "IO".elev[3].jinggao.LC := "INPUT"."3号梯光幕信号";
       "IO".elev[3].jinggao.REP := "INPUT"."3号梯检修信号";

       "IO".elev[3].bt_limit.bottom1 := "INPUT"."3号梯下端站第1限位";
       "IO".elev[3].bt_limit.bottom2 := "INPUT"."3号梯下端站第2限位";
       "IO".elev[3].bt_limit.top1 := "INPUT"."3号梯上端站第1限位";
       "IO".elev[3].bt_limit.top2 := "INPUT"."3号梯上端站第2限位";

       "IO".elev[3].zhongliang := "INPUT"."3号梯当前载重量";
   END_REGION
   REGION 4号梯INPUT
       "IO".elev[4].ele_in_button[1].state := "INPUT"."4号梯轿内选层按钮1";
       "IO".elev[4].ele_in_button[2].state := "INPUT"."4号梯轿内选层按钮2";
       "IO".elev[4].ele_in_button[3].state := "INPUT"."4号梯轿内选层按钮3";
       "IO".elev[4].ele_in_button[4].state := "INPUT"."4号梯轿内选层按钮4";
       "IO".elev[4].ele_in_button[5].state := "INPUT"."4号梯轿内选层按钮5";
       "IO".elev[4].ele_in_button[6].state := "INPUT"."4号梯轿内选层按钮6";
       "IO".elev[4].ele_in_button[7].state := "INPUT"."4号梯轿内选层按钮7";
       "IO".elev[4].ele_in_button[8].state := "INPUT"."4号梯轿内选层按钮8";
       "IO".elev[4].ele_in_button[9].state := "INPUT"."4号梯轿内选层按钮9";
       "IO".elev[4].ele_in_button[10].state := "INPUT"."4号梯轿内选层按钮10";

       "IO".elev[4].door_open.state := "INPUT"."4号梯轿内开门按钮";
       "IO".elev[4].btn_close.state := "INPUT"."4号梯轿内关门按钮";

       "IO".elev[4].door_Lock := "INPUT"."4号梯轿厢门锁信号";
       "IO".elev[4].floor_Lock[1] := "INPUT"."4号梯1楼层门锁信号";
       "IO".elev[4].floor_Lock[2] := "INPUT"."4号梯2楼层门锁信号";
       "IO".elev[4].floor_Lock[3] := "INPUT"."4号梯3楼层门锁信号";
       "IO".elev[4].floor_Lock[4] := "INPUT"."4号梯4楼层门锁信号";
       "IO".elev[4].floor_Lock[5] := "INPUT"."4号梯5楼层门锁信号";
       "IO".elev[4].floor_Lock[6] := "INPUT"."4号梯6楼层门锁信号";
       "IO".elev[4].floor_Lock[7] := "INPUT"."4号梯7楼层门锁信号";
       "IO".elev[4].floor_Lock[8] := "INPUT"."4号梯8楼层门锁信号";
       "IO".elev[4].floor_Lock[9] := "INPUT"."4号梯9楼层门锁信号";
       "IO".elev[4].floor_Lock[10] := "INPUT"."4号梯10楼层门锁信号";

       "IO".elev[4].button_out[1, 1].state := "INPUT"."4号梯1层上行呼梯按钮";
       "IO".elev[4].button_out[1, 2].state := "INPUT"."4号梯2层上行呼梯按钮";
       "IO".elev[4].button_out[1, 3].state := "INPUT"."4号梯3层上行呼梯按钮";
       "IO".elev[4].button_out[1, 4].state := "INPUT"."4号梯4层上行呼梯按钮";
       "IO".elev[4].button_out[1, 5].state := "INPUT"."4号梯5层上行呼梯按钮";
       "IO".elev[4].button_out[1, 6].state := "INPUT"."4号梯6层上行呼梯按钮";
       "IO".elev[4].button_out[1, 7].state := "INPUT"."4号梯7层上行呼梯按钮";
       "IO".elev[4].button_out[1, 8].state := "INPUT"."4号梯8层上行呼梯按钮";
       "IO".elev[4].button_out[1, 9].state := "INPUT"."4号梯9层上行呼梯按钮";

       "IO".elev[4].button_out[2, 2].state := "INPUT"."4号梯2层下行呼梯按钮";
       "IO".elev[4].button_out[2, 3].state := "INPUT"."4号梯3层下行呼梯按钮";
       "IO".elev[4].button_out[2, 4].state := "INPUT"."4号梯4层下行呼梯按钮";
       "IO".elev[4].button_out[2, 5].state := "INPUT"."4号梯5层下行呼梯按钮";
       "IO".elev[4].button_out[2, 6].state := "INPUT"."4号梯6层下行呼梯按钮";
       "IO".elev[4].button_out[2, 7].state := "INPUT"."4号梯7层下行呼梯按钮";
       "IO".elev[4].button_out[2, 8].state := "INPUT"."4号梯8层下行呼梯按钮";
       "IO".elev[4].button_out[2, 9].state := "INPUT"."4号梯9层下行呼梯按钮";
       "IO".elev[4].button_out[2, 10].state := "INPUT"."4号梯10层下行呼梯按钮";

       "IO".elev[4].door_inplace.open := "INPUT"."4号梯开门到位";
       "IO".elev[4].door_inplace.close := "INPUT"."4号梯关门到位";

       "IO".elev[4].direction.up := "INPUT"."4号梯上平层信号";
       "IO".elev[4].direction.down := "INPUT"."4号梯下平层信号";

       "IO".elev[4].jinggao.LC := "INPUT"."4号梯光幕信号";
       "IO".elev[4].jinggao.REP := "INPUT"."4号梯检修信号";

       "IO".elev[4].bt_limit.bottom1 := "INPUT"."4号梯下端站第1限位";
       "IO".elev[4].bt_limit.bottom2 := "INPUT"."4号梯下端站第2限位";
       "IO".elev[4].bt_limit.top1 := "INPUT"."4号梯上端站第1限位";
       "IO".elev[4].bt_limit.top2 := "INPUT"."4号梯上端站第2限位";

       "IO".elev[4].zhongliang := "INPUT"."4号梯当前载重量";
   END_REGION
   REGION 5号梯INPUT
       "IO".elev[5].ele_in_button[1].state := "INPUT"."5号梯轿内选层按钮1";
       "IO".elev[5].ele_in_button[2].state := "INPUT"."5号梯轿内选层按钮2";
       "IO".elev[5].ele_in_button[3].state := "INPUT"."5号梯轿内选层按钮3";
       "IO".elev[5].ele_in_button[4].state := "INPUT"."5号梯轿内选层按钮5";
       "IO".elev[5].ele_in_button[5].state := "INPUT"."5号梯轿内选层按钮5";
       "IO".elev[5].ele_in_button[6].state := "INPUT"."5号梯轿内选层按钮6";
       "IO".elev[5].ele_in_button[7].state := "INPUT"."5号梯轿内选层按钮7";
       "IO".elev[5].ele_in_button[8].state := "INPUT"."5号梯轿内选层按钮8";
       "IO".elev[5].ele_in_button[9].state := "INPUT"."5号梯轿内选层按钮9";
       "IO".elev[5].ele_in_button[10].state := "INPUT"."5号梯轿内选层按钮10";

       "IO".elev[5].door_open.state := "INPUT"."5号梯轿内开门按钮";
       "IO".elev[5].btn_close.state := "INPUT"."5号梯轿内关门按钮";

       "IO".elev[5].door_Lock := "INPUT"."5号梯轿厢门锁信号";
       "IO".elev[5].floor_Lock[1] := "INPUT"."5号梯1楼层门锁信号";
       "IO".elev[5].floor_Lock[2] := "INPUT"."5号梯2楼层门锁信号";
       "IO".elev[5].floor_Lock[3] := "INPUT"."5号梯3楼层门锁信号";
       "IO".elev[5].floor_Lock[4] := "INPUT"."5号梯4楼层门锁信号";
       "IO".elev[5].floor_Lock[5] := "INPUT"."5号梯5楼层门锁信号";
       "IO".elev[5].floor_Lock[6] := "INPUT"."5号梯6楼层门锁信号";
       "IO".elev[5].floor_Lock[7] := "INPUT"."5号梯7楼层门锁信号";
       "IO".elev[5].floor_Lock[8] := "INPUT"."5号梯8楼层门锁信号";
       "IO".elev[5].floor_Lock[9] := "INPUT"."5号梯9楼层门锁信号";
       "IO".elev[5].floor_Lock[10] := "INPUT"."5号梯10楼层门锁信号";

       "IO".elev[5].button_out[1, 1].state := "INPUT"."5号梯1层上行呼梯按钮";
       "IO".elev[5].button_out[1, 2].state := "INPUT"."5号梯2层上行呼梯按钮";
       "IO".elev[5].button_out[1, 3].state := "INPUT"."5号梯3层上行呼梯按钮";
       "IO".elev[5].button_out[1, 4].state := "INPUT"."5号梯4层上行呼梯按钮";
       "IO".elev[5].button_out[1, 5].state := "INPUT"."5号梯5层上行呼梯按钮";
       "IO".elev[5].button_out[1, 6].state := "INPUT"."5号梯6层上行呼梯按钮";
       "IO".elev[5].button_out[1, 7].state := "INPUT"."5号梯7层上行呼梯按钮";
       "IO".elev[5].button_out[1, 8].state := "INPUT"."5号梯8层上行呼梯按钮";
       "IO".elev[5].button_out[1, 9].state := "INPUT"."5号梯9层上行呼梯按钮";

       "IO".elev[5].button_out[2, 2].state := "INPUT"."5号梯2层下行呼梯按钮";
       "IO".elev[5].button_out[2, 3].state := "INPUT"."5号梯3层下行呼梯按钮";
       "IO".elev[5].button_out[2, 4].state := "INPUT"."5号梯4层下行呼梯按钮";
       "IO".elev[5].button_out[2, 5].state := "INPUT"."5号梯5层下行呼梯按钮";
       "IO".elev[5].button_out[2, 6].state := "INPUT"."5号梯6层下行呼梯按钮";
       "IO".elev[5].button_out[2, 7].state := "INPUT"."5号梯7层下行呼梯按钮";
       "IO".elev[5].button_out[2, 8].state := "INPUT"."5号梯8层下行呼梯按钮";
       "IO".elev[5].button_out[2, 9].state := "INPUT"."5号梯9层下行呼梯按钮";
       "IO".elev[5].button_out[2, 10].state := "INPUT"."5号梯10层下行呼梯按钮";

       "IO".elev[5].door_inplace.open := "INPUT"."5号梯开门到位";
       "IO".elev[5].door_inplace.close := "INPUT"."5号梯关门到位";

       "IO".elev[5].direction.up := "INPUT"."5号梯上平层信号";
       "IO".elev[5].direction.down := "INPUT"."5号梯下平层信号";

       "IO".elev[5].jinggao.LC := "INPUT"."5号梯光幕信号";
       "IO".elev[5].jinggao.REP := "INPUT"."5号梯检修信号";

       "IO".elev[5].bt_limit.bottom1 := "INPUT"."5号梯下端站第1限位";
       "IO".elev[5].bt_limit.bottom2 := "INPUT"."5号梯下端站第2限位";
       "IO".elev[5].bt_limit.top1 := "INPUT"."5号梯上端站第1限位";
       "IO".elev[5].bt_limit.top2 := "INPUT"."5号梯上端站第2限位";

       "IO".elev[5].zhongliang := "INPUT"."5号梯当前载重量";
   END_REGION
   REGION 6号梯INPUT
       "IO".elev[6].ele_in_button[1].state := "INPUT"."6号梯轿内选层按钮1";
       "IO".elev[6].ele_in_button[2].state := "INPUT"."6号梯轿内选层按钮2";
       "IO".elev[6].ele_in_button[3].state := "INPUT"."6号梯轿内选层按钮3";
       "IO".elev[6].ele_in_button[4].state := "INPUT"."6号梯轿内选层按钮6";
       "IO".elev[6].ele_in_button[5].state := "INPUT"."6号梯轿内选层按钮6";
       "IO".elev[6].ele_in_button[6].state := "INPUT"."6号梯轿内选层按钮6";
       "IO".elev[6].ele_in_button[7].state := "INPUT"."6号梯轿内选层按钮7";
       "IO".elev[6].ele_in_button[8].state := "INPUT"."6号梯轿内选层按钮8";
       "IO".elev[6].ele_in_button[9].state := "INPUT"."6号梯轿内选层按钮9";
       "IO".elev[6].ele_in_button[10].state := "INPUT"."6号梯轿内选层按钮10";

       "IO".elev[6].door_open.state := "INPUT"."6号梯轿内开门按钮";
       "IO".elev[6].btn_close.state := "INPUT"."6号梯轿内关门按钮";

       "IO".elev[6].door_Lock := "INPUT"."6号梯轿厢门锁信号";
       "IO".elev[6].floor_Lock[1] := "INPUT"."6号梯1楼层门锁信号";
       "IO".elev[6].floor_Lock[2] := "INPUT"."6号梯2楼层门锁信号";
       "IO".elev[6].floor_Lock[3] := "INPUT"."6号梯3楼层门锁信号";
       "IO".elev[6].floor_Lock[4] := "INPUT"."6号梯4楼层门锁信号";
       "IO".elev[6].floor_Lock[5] := "INPUT"."6号梯5楼层门锁信号";
       "IO".elev[6].floor_Lock[6] := "INPUT"."6号梯6楼层门锁信号";
       "IO".elev[6].floor_Lock[7] := "INPUT"."6号梯7楼层门锁信号";
       "IO".elev[6].floor_Lock[8] := "INPUT"."6号梯8楼层门锁信号";
       "IO".elev[6].floor_Lock[9] := "INPUT"."6号梯9楼层门锁信号";
       "IO".elev[6].floor_Lock[10] := "INPUT"."6号梯10楼层门锁信号";

       "IO".elev[6].button_out[1, 1].state := "INPUT"."6号梯1层上行呼梯按钮";
       "IO".elev[6].button_out[1, 2].state := "INPUT"."6号梯2层上行呼梯按钮";
       "IO".elev[6].button_out[1, 3].state := "INPUT"."6号梯3层上行呼梯按钮";
       "IO".elev[6].button_out[1, 4].state := "INPUT"."6号梯4层上行呼梯按钮";
       "IO".elev[6].button_out[1, 5].state := "INPUT"."6号梯5层上行呼梯按钮";
       "IO".elev[6].button_out[1, 6].state := "INPUT"."6号梯6层上行呼梯按钮";
       "IO".elev[6].button_out[1, 7].state := "INPUT"."6号梯7层上行呼梯按钮";
       "IO".elev[6].button_out[1, 8].state := "INPUT"."6号梯8层上行呼梯按钮";
       "IO".elev[6].button_out[1, 9].state := "INPUT"."6号梯9层上行呼梯按钮";

       "IO".elev[6].button_out[2, 2].state := "INPUT"."6号梯2层下行呼梯按钮";
       "IO".elev[6].button_out[2, 3].state := "INPUT"."6号梯3层下行呼梯按钮";
       "IO".elev[6].button_out[2, 4].state := "INPUT"."6号梯4层下行呼梯按钮";
       "IO".elev[6].button_out[2, 5].state := "INPUT"."6号梯5层下行呼梯按钮";
       "IO".elev[6].button_out[2, 6].state := "INPUT"."6号梯6层下行呼梯按钮";
       "IO".elev[6].button_out[2, 7].state := "INPUT"."6号梯7层下行呼梯按钮";
       "IO".elev[6].button_out[2, 8].state := "INPUT"."6号梯8层下行呼梯按钮";
       "IO".elev[6].button_out[2, 9].state := "INPUT"."6号梯9层下行呼梯按钮";
       "IO".elev[6].button_out[2, 10].state := "INPUT"."6号梯10层下行呼梯按钮";

       "IO".elev[6].door_inplace.open := "INPUT"."6号梯开门到位";
       "IO".elev[6].door_inplace.close := "INPUT"."6号梯关门到位";

       "IO".elev[6].direction.up := "INPUT"."6号梯上平层信号";
       "IO".elev[6].direction.down := "INPUT"."6号梯下平层信号";

       "IO".elev[6].jinggao.LC := "INPUT"."6号梯光幕信号";
       "IO".elev[6].jinggao.REP := "INPUT"."6号梯检修信号";

       "IO".elev[6].bt_limit.bottom1 := "INPUT"."6号梯下端站第1限位";
       "IO".elev[6].bt_limit.bottom2 := "INPUT"."6号梯下端站第2限位";
       "IO".elev[6].bt_limit.top1 := "INPUT"."6号梯上端站第1限位";
       "IO".elev[6].bt_limit.top2 := "INPUT"."6号梯上端站第2限位";

       "IO".elev[6].zhongliang := "INPUT"."6号梯当前载重量";
   END_REGION
   //************************************************************************************************************************//
   //***********************************************OUTPUT*******************************************************************//
   REGION 公共部分
       "OUTPUT".准备就绪信号 := "IO".plc_ready;

   END_REGION
   REGION 1号梯OUTPUT
       "OUTPUT"."1号梯1层按钮指示灯" := "IO".elev[1].ele_in_button[1].light;
       "OUTPUT"."1号梯2层按钮指示灯" := "IO".elev[1].ele_in_button[2].light;
       "OUTPUT"."1号梯3层按钮指示灯" := "IO".elev[1].ele_in_button[3].light;
       "OUTPUT"."1号梯4层按钮指示灯" := "IO".elev[1].ele_in_button[4].light;
       "OUTPUT"."1号梯5层按钮指示灯" := "IO".elev[1].ele_in_button[5].light;
       "OUTPUT"."1号梯6层按钮指示灯" := "IO".elev[1].ele_in_button[6].light;
       "OUTPUT"."1号梯7层按钮指示灯" := "IO".elev[1].ele_in_button[7].light;
       "OUTPUT"."1号梯8层按钮指示灯" := "IO".elev[1].ele_in_button[8].light;
       "OUTPUT"."1号梯9层按钮指示灯" := "IO".elev[1].ele_in_button[9].light;
       "OUTPUT"."1号梯10层按钮指示灯" := "IO".elev[1].ele_in_button[10].light;

       "OUTPUT"."1号梯1层上行呼梯按钮指示灯" := "IO".elev[1].button_out[1, 1].light;
       "OUTPUT"."1号梯2层上行呼梯按钮指示灯" := "IO".elev[1].button_out[1, 2].light;
       "OUTPUT"."1号梯3层上行呼梯按钮指示灯" := "IO".elev[1].button_out[1, 3].light;
       "OUTPUT"."1号梯4层上行呼梯按钮指示灯" := "IO".elev[1].button_out[1, 4].light;
       "OUTPUT"."1号梯5层上行呼梯按钮指示灯" := "IO".elev[1].button_out[1, 5].light;
       "OUTPUT"."1号梯6层上行呼梯按钮指示灯" := "IO".elev[1].button_out[1, 6].light;
       "OUTPUT"."1号梯7层上行呼梯按钮指示灯" := "IO".elev[1].button_out[1, 7].light;
       "OUTPUT"."1号梯8层上行呼梯按钮指示灯" := "IO".elev[1].button_out[1, 8].light;
       "OUTPUT"."1号梯9层上行呼梯按钮指示灯" := "IO".elev[1].button_out[1, 9].light;

       "OUTPUT"."1号梯2层下行呼梯按钮指示灯" := "IO".elev[1].button_out[2, 2].light;
       "OUTPUT"."1号梯3层下行呼梯按钮指示灯" := "IO".elev[1].button_out[2, 3].light;
       "OUTPUT"."1号梯4层下行呼梯按钮指示灯" := "IO".elev[1].button_out[2, 4].light;
       "OUTPUT"."1号梯5层下行呼梯按钮指示灯" := "IO".elev[1].button_out[2, 5].light;
       "OUTPUT"."1号梯6层下行呼梯按钮指示灯" := "IO".elev[1].button_out[2, 6].light;
       "OUTPUT"."1号梯7层下行呼梯按钮指示灯" := "IO".elev[1].button_out[2, 7].light;
       "OUTPUT"."1号梯8层下行呼梯按钮指示灯" := "IO".elev[1].button_out[2, 8].light;
       "OUTPUT"."1号梯9层下行呼梯按钮指示灯" := "IO".elev[1].button_out[2, 9].light;
       "OUTPUT"."1号梯10层下行呼梯按钮指示灯" := "IO".elev[1].button_out[2, 10].light;

       "OUTPUT"."1号梯LEDa" := "IO".elev[1].smg[1, 1];
       "OUTPUT"."1号梯LEDb" := "IO".elev[1].smg[1, 2];
       "OUTPUT"."1号梯LEDc" := "IO".elev[1].smg[1, 3];
       "OUTPUT"."1号梯LEDd" := "IO".elev[1].smg[1, 4];
       "OUTPUT"."1号梯LEDe" := "IO".elev[1].smg[1, 5];
       "OUTPUT"."1号梯LEDf" := "IO".elev[1].smg[1, 6];
       "OUTPUT"."1号梯LEDg" := "IO".elev[1].smg[1, 7];
       "OUTPUT"."1号梯LEDh" := "IO".elev[1].smg[2, 1];
       "OUTPUT"."1号梯LEDi" := "IO".elev[1].smg[2, 2];
       "OUTPUT"."1号梯LEDj" := "IO".elev[1].smg[2, 3];
       "OUTPUT"."1号梯LEDk" := "IO".elev[1].smg[2, 4];
       "OUTPUT"."1号梯LEDl" := "IO".elev[1].smg[2, 5];
       "OUTPUT"."1号梯LEDm" := "IO".elev[1].smg[2, 6];
       "OUTPUT"."1号梯LEDn" := "IO".elev[1].smg[2, 7];

       "OUTPUT"."1号梯风扇指示" := "IO".elev[1].display.fan;
       "OUTPUT"."1号梯故障指示" := "IO".elev[1].display.error;
       "OUTPUT"."1号梯满载指示" := "IO".elev[1].display.full;
       "OUTPUT"."1号梯照明指示" := "IO".elev[1].display.light;

       "OUTPUT"."1号梯上行指示" := "IO".elev[1].run_disp.up;
       "OUTPUT"."1号梯下行指示" := "IO".elev[1].run_disp.dowm;

       "OUTPUT"."1号梯1级减速制动" := "IO".elev[1].Brake.B1;
       "OUTPUT"."1号梯2级减速制动" := "IO".elev[1].Brake.B2;
       "OUTPUT"."1号梯3级减速制动" := "IO".elev[1].Brake.B3;

       "OUTPUT"."1号梯高速接触器" := "IO".elev[1].ele_speed.H;
       "OUTPUT"."1号梯低速接触器" := "IO".elev[1].ele_speed.L;

       "OUTPUT"."1号梯电机启动信号" := "IO".elev[1].run_enable;
       "OUTPUT"."1号梯上行接触器" := "IO".elev[1].run_contactor.up;
       "OUTPUT"."1号梯下行接触器" := "IO".elev[1].run_contactor.dowm;

       "OUTPUT"."1号梯开门继电器" := "IO".elev[1].door_jdq.open;
       "OUTPUT"."1号梯关门继电器" := "IO".elev[1].door_jdq.close;
   END_REGION
   REGION 2号梯OUTPUT
       "OUTPUT"."2号梯1层按钮指示灯" := "IO".elev[2].ele_in_button[1].light;
       "OUTPUT"."2号梯2层按钮指示灯" := "IO".elev[2].ele_in_button[2].light;
       "OUTPUT"."2号梯3层按钮指示灯" := "IO".elev[2].ele_in_button[3].light;
       "OUTPUT"."2号梯4层按钮指示灯" := "IO".elev[2].ele_in_button[4].light;
       "OUTPUT"."2号梯5层按钮指示灯" := "IO".elev[2].ele_in_button[5].light;
       "OUTPUT"."2号梯6层按钮指示灯" := "IO".elev[2].ele_in_button[6].light;
       "OUTPUT"."2号梯7层按钮指示灯" := "IO".elev[2].ele_in_button[7].light;
       "OUTPUT"."2号梯8层按钮指示灯" := "IO".elev[2].ele_in_button[8].light;
       "OUTPUT"."2号梯9层按钮指示灯" := "IO".elev[2].ele_in_button[9].light;
       "OUTPUT"."2号梯10层按钮指示灯" := "IO".elev[2].ele_in_button[10].light;

       "OUTPUT"."2号梯1层上行呼梯按钮指示灯" := "IO".elev[2].button_out[1, 1].light;
       "OUTPUT"."2号梯2层上行呼梯按钮指示灯" := "IO".elev[2].button_out[1, 2].light;
       "OUTPUT"."2号梯3层上行呼梯按钮指示灯" := "IO".elev[2].button_out[1, 3].light;
       "OUTPUT"."2号梯4层上行呼梯按钮指示灯" := "IO".elev[2].button_out[1, 4].light;
       "OUTPUT"."2号梯5层上行呼梯按钮指示灯" := "IO".elev[2].button_out[1, 5].light;
       "OUTPUT"."2号梯6层上行呼梯按钮指示灯" := "IO".elev[2].button_out[1, 6].light;
       "OUTPUT"."2号梯7层上行呼梯按钮指示灯" := "IO".elev[2].button_out[1, 7].light;
       "OUTPUT"."2号梯8层上行呼梯按钮指示灯" := "IO".elev[2].button_out[1, 8].light;
       "OUTPUT"."2号梯9层上行呼梯按钮指示灯" := "IO".elev[2].button_out[1, 9].light;

       "OUTPUT"."2号梯2层下行呼梯按钮指示灯" := "IO".elev[2].button_out[2, 2].light;
       "OUTPUT"."2号梯3层下行呼梯按钮指示灯" := "IO".elev[2].button_out[2, 3].light;
       "OUTPUT"."2号梯4层下行呼梯按钮指示灯" := "IO".elev[2].button_out[2, 4].light;
       "OUTPUT"."2号梯5层下行呼梯按钮指示灯" := "IO".elev[2].button_out[2, 5].light;
       "OUTPUT"."2号梯6层下行呼梯按钮指示灯" := "IO".elev[2].button_out[2, 6].light;
       "OUTPUT"."2号梯7层下行呼梯按钮指示灯" := "IO".elev[2].button_out[2, 7].light;
       "OUTPUT"."2号梯8层下行呼梯按钮指示灯" := "IO".elev[2].button_out[2, 8].light;
       "OUTPUT"."2号梯9层下行呼梯按钮指示灯" := "IO".elev[2].button_out[2, 9].light;
       "OUTPUT"."2号梯10层下行呼梯按钮指示灯" := "IO".elev[2].button_out[2, 10].light;

       "OUTPUT"."2号梯LEDa" := "IO".elev[2].smg[1, 1];
       "OUTPUT"."2号梯LEDb" := "IO".elev[2].smg[1, 2];
       "OUTPUT"."2号梯LEDc" := "IO".elev[2].smg[1, 3];
       "OUTPUT"."2号梯LEDd" := "IO".elev[2].smg[1, 4];
       "OUTPUT"."2号梯LEDe" := "IO".elev[2].smg[1, 5];
       "OUTPUT"."2号梯LEDf" := "IO".elev[2].smg[1, 6];
       "OUTPUT"."2号梯LEDg" := "IO".elev[2].smg[1, 7];
       "OUTPUT"."2号梯LEDh" := "IO".elev[2].smg[2, 1];
       "OUTPUT"."2号梯LEDi" := "IO".elev[2].smg[2, 2];
       "OUTPUT"."2号梯LEDj" := "IO".elev[2].smg[2, 3];
       "OUTPUT"."2号梯LEDk" := "IO".elev[2].smg[2, 4];
       "OUTPUT"."2号梯LEDl" := "IO".elev[2].smg[2, 5];
       "OUTPUT"."2号梯LEDm" := "IO".elev[2].smg[2, 6];
       "OUTPUT"."2号梯LEDn" := "IO".elev[2].smg[2, 7];

       "OUTPUT"."2号梯风扇指示" := "IO".elev[2].display.fan;
       "OUTPUT"."2号梯故障指示" := "IO".elev[2].display.error;
       "OUTPUT"."2号梯满载指示" := "IO".elev[2].display.full;
       "OUTPUT"."2号梯照明指示" := "IO".elev[2].display.light;

       "OUTPUT"."2号梯上行指示" := "IO".elev[2].run_disp.up;
       "OUTPUT"."2号梯下行指示" := "IO".elev[2].run_disp.dowm;

       "OUTPUT"."2号梯1级减速制动" := "IO".elev[2].Brake.B1;
       "OUTPUT"."2号梯2级减速制动" := "IO".elev[2].Brake.B2;
       "OUTPUT"."2号梯3级减速制动" := "IO".elev[2].Brake.B3;

       "OUTPUT"."2号梯高速接触器" := "IO".elev[2].ele_speed.H;
       "OUTPUT"."2号梯低速接触器" := "IO".elev[2].ele_speed.L;

       "OUTPUT"."2号梯电机启动信号" := "IO".elev[2].run_enable;
       "OUTPUT"."2号梯上行接触器" := "IO".elev[2].run_contactor.up;
       "OUTPUT"."2号梯下行接触器" := "IO".elev[2].run_contactor.dowm;

       "OUTPUT"."2号梯开门继电器" := "IO".elev[2].door_jdq.open;
       "OUTPUT"."2号梯关门继电器" := "IO".elev[2].door_jdq.close;
   END_REGION
   REGION 3号梯OUTPUT
       "OUTPUT"."3号梯1层按钮指示灯" := "IO".elev[3].ele_in_button[1].light;
       "OUTPUT"."3号梯2层按钮指示灯" := "IO".elev[3].ele_in_button[2].light;
       "OUTPUT"."3号梯3层按钮指示灯" := "IO".elev[3].ele_in_button[3].light;
       "OUTPUT"."3号梯4层按钮指示灯" := "IO".elev[3].ele_in_button[4].light;
       "OUTPUT"."3号梯5层按钮指示灯" := "IO".elev[3].ele_in_button[5].light;
       "OUTPUT"."3号梯6层按钮指示灯" := "IO".elev[3].ele_in_button[6].light;
       "OUTPUT"."3号梯7层按钮指示灯" := "IO".elev[3].ele_in_button[7].light;
       "OUTPUT"."3号梯8层按钮指示灯" := "IO".elev[3].ele_in_button[8].light;
       "OUTPUT"."3号梯9层按钮指示灯" := "IO".elev[3].ele_in_button[9].light;
       "OUTPUT"."3号梯10层按钮指示灯" := "IO".elev[3].ele_in_button[10].light;

       "OUTPUT"."3号梯1层上行呼梯按钮指示灯" := "IO".elev[3].button_out[1, 1].light;
       "OUTPUT"."3号梯2层上行呼梯按钮指示灯" := "IO".elev[3].button_out[1, 2].light;
       "OUTPUT"."3号梯3层上行呼梯按钮指示灯" := "IO".elev[3].button_out[1, 3].light;
       "OUTPUT"."3号梯4层上行呼梯按钮指示灯" := "IO".elev[3].button_out[1, 4].light;
       "OUTPUT"."3号梯5层上行呼梯按钮指示灯" := "IO".elev[3].button_out[1, 5].light;
       "OUTPUT"."3号梯6层上行呼梯按钮指示灯" := "IO".elev[3].button_out[1, 6].light;
       "OUTPUT"."3号梯7层上行呼梯按钮指示灯" := "IO".elev[3].button_out[1, 7].light;
       "OUTPUT"."3号梯8层上行呼梯按钮指示灯" := "IO".elev[3].button_out[1, 8].light;
       "OUTPUT"."3号梯9层上行呼梯按钮指示灯" := "IO".elev[3].button_out[1, 9].light;

       "OUTPUT"."3号梯2层下行呼梯按钮指示灯" := "IO".elev[3].button_out[2, 2].light;
       "OUTPUT"."3号梯3层下行呼梯按钮指示灯" := "IO".elev[3].button_out[2, 3].light;
       "OUTPUT"."3号梯4层下行呼梯按钮指示灯" := "IO".elev[3].button_out[2, 4].light;
       "OUTPUT"."3号梯5层下行呼梯按钮指示灯" := "IO".elev[3].button_out[2, 5].light;
       "OUTPUT"."3号梯6层下行呼梯按钮指示灯" := "IO".elev[3].button_out[2, 6].light;
       "OUTPUT"."3号梯7层下行呼梯按钮指示灯" := "IO".elev[3].button_out[2, 7].light;
       "OUTPUT"."3号梯8层下行呼梯按钮指示灯" := "IO".elev[3].button_out[2, 8].light;
       "OUTPUT"."3号梯9层下行呼梯按钮指示灯" := "IO".elev[3].button_out[2, 9].light;
       "OUTPUT"."3号梯10层下行呼梯按钮指示灯" := "IO".elev[3].button_out[2, 10].light;

       "OUTPUT"."3号梯LEDa" := "IO".elev[3].smg[1, 1];
       "OUTPUT"."3号梯LEDb" := "IO".elev[3].smg[1, 2];
       "OUTPUT"."3号梯LEDc" := "IO".elev[3].smg[1, 3];
       "OUTPUT"."3号梯LEDd" := "IO".elev[3].smg[1, 4];
       "OUTPUT"."3号梯LEDe" := "IO".elev[3].smg[1, 5];
       "OUTPUT"."3号梯LEDf" := "IO".elev[3].smg[1, 6];
       "OUTPUT"."3号梯LEDg" := "IO".elev[3].smg[1, 7];
       "OUTPUT"."3号梯LEDh" := "IO".elev[3].smg[2, 1];
       "OUTPUT"."3号梯LEDi" := "IO".elev[3].smg[2, 2];
       "OUTPUT"."3号梯LEDj" := "IO".elev[3].smg[2, 3];
       "OUTPUT"."3号梯LEDk" := "IO".elev[3].smg[2, 4];
       "OUTPUT"."3号梯LEDl" := "IO".elev[3].smg[2, 5];
       "OUTPUT"."3号梯LEDm" := "IO".elev[3].smg[2, 6];
       "OUTPUT"."3号梯LEDn" := "IO".elev[3].smg[2, 7];

       "OUTPUT"."3号梯风扇指示" := "IO".elev[3].display.fan;
       "OUTPUT"."3号梯故障指示" := "IO".elev[3].display.error;
       "OUTPUT"."3号梯满载指示" := "IO".elev[3].display.full;
       "OUTPUT"."3号梯照明指示" := "IO".elev[3].display.light;

       "OUTPUT"."3号梯上行指示" := "IO".elev[3].run_disp.up;
       "OUTPUT"."3号梯下行指示" := "IO".elev[3].run_disp.dowm;

       "OUTPUT"."3号梯1级减速制动" := "IO".elev[3].Brake.B1;
       "OUTPUT"."3号梯2级减速制动" := "IO".elev[3].Brake.B2;
       "OUTPUT"."3号梯3级减速制动" := "IO".elev[3].Brake.B3;

       "OUTPUT"."3号梯高速接触器" := "IO".elev[3].ele_speed.H;
       "OUTPUT"."3号梯低速接触器" := "IO".elev[3].ele_speed.L;

       "OUTPUT"."3号梯电机启动信号" := "IO".elev[3].run_enable;
       "OUTPUT"."3号梯上行接触器" := "IO".elev[3].run_contactor.up;
       "OUTPUT"."3号梯下行接触器" := "IO".elev[3].run_contactor.dowm;

       "OUTPUT"."3号梯开门继电器" := "IO".elev[3].door_jdq.open;
       "OUTPUT"."3号梯关门继电器" := "IO".elev[3].door_jdq.close;
   END_REGION
   REGION 4号梯OUTPUT
       "OUTPUT"."4号梯1层按钮指示灯" := "IO".elev[4].ele_in_button[1].light;
       "OUTPUT"."4号梯2层按钮指示灯" := "IO".elev[4].ele_in_button[2].light;
       "OUTPUT"."4号梯3层按钮指示灯" := "IO".elev[4].ele_in_button[3].light;
       "OUTPUT"."4号梯4层按钮指示灯" := "IO".elev[4].ele_in_button[4].light;
       "OUTPUT"."4号梯5层按钮指示灯" := "IO".elev[4].ele_in_button[5].light;
       "OUTPUT"."4号梯6层按钮指示灯" := "IO".elev[4].ele_in_button[6].light;
       "OUTPUT"."4号梯7层按钮指示灯" := "IO".elev[4].ele_in_button[7].light;
       "OUTPUT"."4号梯8层按钮指示灯" := "IO".elev[4].ele_in_button[8].light;
       "OUTPUT"."4号梯9层按钮指示灯" := "IO".elev[4].ele_in_button[9].light;
       "OUTPUT"."4号梯10层按钮指示灯" := "IO".elev[4].ele_in_button[10].light;

       "OUTPUT"."4号梯1层上行呼梯按钮指示灯" := "IO".elev[4].button_out[1, 1].light;
       "OUTPUT"."4号梯2层上行呼梯按钮指示灯" := "IO".elev[4].button_out[1, 2].light;
       "OUTPUT"."4号梯3层上行呼梯按钮指示灯" := "IO".elev[4].button_out[1, 3].light;
       "OUTPUT"."4号梯4层上行呼梯按钮指示灯" := "IO".elev[4].button_out[1, 4].light;
       "OUTPUT"."4号梯5层上行呼梯按钮指示灯" := "IO".elev[4].button_out[1, 5].light;
       "OUTPUT"."4号梯6层上行呼梯按钮指示灯" := "IO".elev[4].button_out[1, 6].light;
       "OUTPUT"."4号梯7层上行呼梯按钮指示灯" := "IO".elev[4].button_out[1, 7].light;
       "OUTPUT"."4号梯8层上行呼梯按钮指示灯" := "IO".elev[4].button_out[1, 8].light;
       "OUTPUT"."4号梯9层上行呼梯按钮指示灯" := "IO".elev[4].button_out[1, 9].light;

       "OUTPUT"."4号梯2层下行呼梯按钮指示灯" := "IO".elev[4].button_out[2, 2].light;
       "OUTPUT"."4号梯3层下行呼梯按钮指示灯" := "IO".elev[4].button_out[2, 3].light;
       "OUTPUT"."4号梯4层下行呼梯按钮指示灯" := "IO".elev[4].button_out[2, 4].light;
       "OUTPUT"."4号梯5层下行呼梯按钮指示灯" := "IO".elev[4].button_out[2, 5].light;
       "OUTPUT"."4号梯6层下行呼梯按钮指示灯" := "IO".elev[4].button_out[2, 6].light;
       "OUTPUT"."4号梯7层下行呼梯按钮指示灯" := "IO".elev[4].button_out[2, 7].light;
       "OUTPUT"."4号梯8层下行呼梯按钮指示灯" := "IO".elev[4].button_out[2, 8].light;
       "OUTPUT"."4号梯9层下行呼梯按钮指示灯" := "IO".elev[4].button_out[2, 9].light;
       "OUTPUT"."4号梯10层下行呼梯按钮指示灯" := "IO".elev[4].button_out[2, 10].light;

       "OUTPUT"."4号梯LEDa" := "IO".elev[4].smg[1, 1];
       "OUTPUT"."4号梯LEDb" := "IO".elev[4].smg[1, 2];
       "OUTPUT"."4号梯LEDc" := "IO".elev[4].smg[1, 3];
       "OUTPUT"."4号梯LEDd" := "IO".elev[4].smg[1, 4];
       "OUTPUT"."4号梯LEDe" := "IO".elev[4].smg[1, 5];
       "OUTPUT"."4号梯LEDf" := "IO".elev[4].smg[1, 6];
       "OUTPUT"."4号梯LEDg" := "IO".elev[4].smg[1, 7];
       "OUTPUT"."4号梯LEDh" := "IO".elev[4].smg[2, 1];
       "OUTPUT"."4号梯LEDi" := "IO".elev[4].smg[2, 2];
       "OUTPUT"."4号梯LEDj" := "IO".elev[4].smg[2, 3];
       "OUTPUT"."4号梯LEDk" := "IO".elev[4].smg[2, 4];
       "OUTPUT"."4号梯LEDl" := "IO".elev[4].smg[2, 5];
       "OUTPUT"."4号梯LEDm" := "IO".elev[4].smg[2, 6];
       "OUTPUT"."4号梯LEDn" := "IO".elev[4].smg[2, 7];

       "OUTPUT"."4号梯风扇指示" := "IO".elev[4].display.fan;
       "OUTPUT"."4号梯故障指示" := "IO".elev[4].display.error;
       "OUTPUT"."4号梯满载指示" := "IO".elev[4].display.full;
       "OUTPUT"."4号梯照明指示" := "IO".elev[4].display.light;

       "OUTPUT"."4号梯上行指示" := "IO".elev[4].run_disp.up;
       "OUTPUT"."4号梯下行指示" := "IO".elev[4].run_disp.dowm;

       "OUTPUT"."4号梯1级减速制动" := "IO".elev[4].Brake.B1;
       "OUTPUT"."4号梯2级减速制动" := "IO".elev[4].Brake.B2;
       "OUTPUT"."4号梯3级减速制动" := "IO".elev[4].Brake.B3;

       "OUTPUT"."4号梯高速接触器" := "IO".elev[4].ele_speed.H;
       "OUTPUT"."4号梯低速接触器" := "IO".elev[4].ele_speed.L;

       "OUTPUT"."4号梯电机启动信号" := "IO".elev[4].run_enable;
       "OUTPUT"."4号梯上行接触器" := "IO".elev[4].run_contactor.up;
       "OUTPUT"."4号梯下行接触器" := "IO".elev[4].run_contactor.dowm;

       "OUTPUT"."4号梯开门继电器" := "IO".elev[4].door_jdq.open;
       "OUTPUT"."4号梯关门继电器" := "IO".elev[4].door_jdq.close;
   END_REGION
   REGION 5号梯OUTPUT
       "OUTPUT"."5号梯1层按钮指示灯" := "IO".elev[5].ele_in_button[1].light;
       "OUTPUT"."5号梯2层按钮指示灯" := "IO".elev[5].ele_in_button[2].light;
       "OUTPUT"."5号梯3层按钮指示灯" := "IO".elev[5].ele_in_button[3].light;
       "OUTPUT"."5号梯4层按钮指示灯" := "IO".elev[5].ele_in_button[4].light;
       "OUTPUT"."5号梯5层按钮指示灯" := "IO".elev[5].ele_in_button[5].light;
       "OUTPUT"."5号梯6层按钮指示灯" := "IO".elev[5].ele_in_button[6].light;
       "OUTPUT"."5号梯7层按钮指示灯" := "IO".elev[5].ele_in_button[7].light;
       "OUTPUT"."5号梯8层按钮指示灯" := "IO".elev[5].ele_in_button[8].light;
       "OUTPUT"."5号梯9层按钮指示灯" := "IO".elev[5].ele_in_button[9].light;
       "OUTPUT"."5号梯10层按钮指示灯" := "IO".elev[5].ele_in_button[10].light;

       "OUTPUT"."5号梯1层上行呼梯按钮指示灯" := "IO".elev[5].button_out[1, 1].light;
       "OUTPUT"."5号梯2层上行呼梯按钮指示灯" := "IO".elev[5].button_out[1, 2].light;
       "OUTPUT"."5号梯3层上行呼梯按钮指示灯" := "IO".elev[5].button_out[1, 3].light;
       "OUTPUT"."5号梯4层上行呼梯按钮指示灯" := "IO".elev[5].button_out[1, 4].light;
       "OUTPUT"."5号梯5层上行呼梯按钮指示灯" := "IO".elev[5].button_out[1, 5].light;
       "OUTPUT"."5号梯6层上行呼梯按钮指示灯" := "IO".elev[5].button_out[1, 6].light;
       "OUTPUT"."5号梯7层上行呼梯按钮指示灯" := "IO".elev[5].button_out[1, 7].light;
       "OUTPUT"."5号梯8层上行呼梯按钮指示灯" := "IO".elev[5].button_out[1, 8].light;
       "OUTPUT"."5号梯9层上行呼梯按钮指示灯" := "IO".elev[5].button_out[1, 9].light;

       "OUTPUT"."5号梯2层下行呼梯按钮指示灯" := "IO".elev[5].button_out[2, 2].light;
       "OUTPUT"."5号梯3层下行呼梯按钮指示灯" := "IO".elev[5].button_out[2, 3].light;
       "OUTPUT"."5号梯4层下行呼梯按钮指示灯" := "IO".elev[5].button_out[2, 4].light;
       "OUTPUT"."5号梯5层下行呼梯按钮指示灯" := "IO".elev[5].button_out[2, 5].light;
       "OUTPUT"."5号梯6层下行呼梯按钮指示灯" := "IO".elev[5].button_out[2, 6].light;
       "OUTPUT"."5号梯7层下行呼梯按钮指示灯" := "IO".elev[5].button_out[2, 7].light;
       "OUTPUT"."5号梯8层下行呼梯按钮指示灯" := "IO".elev[5].button_out[2, 8].light;
       "OUTPUT"."5号梯9层下行呼梯按钮指示灯" := "IO".elev[5].button_out[2, 9].light;
       "OUTPUT"."5号梯10层下行呼梯按钮指示灯" := "IO".elev[5].button_out[2, 10].light;

       "OUTPUT"."5号梯LEDa" := "IO".elev[5].smg[1, 1];
       "OUTPUT"."5号梯LEDb" := "IO".elev[5].smg[1, 2];
       "OUTPUT"."5号梯LEDc" := "IO".elev[5].smg[1, 3];
       "OUTPUT"."5号梯LEDd" := "IO".elev[5].smg[1, 4];
       "OUTPUT"."5号梯LEDe" := "IO".elev[5].smg[1, 5];
       "OUTPUT"."5号梯LEDf" := "IO".elev[5].smg[1, 6];
       "OUTPUT"."5号梯LEDg" := "IO".elev[5].smg[1, 7];
       "OUTPUT"."5号梯LEDh" := "IO".elev[5].smg[2, 1];
       "OUTPUT"."5号梯LEDi" := "IO".elev[5].smg[2, 2];
       "OUTPUT"."5号梯LEDj" := "IO".elev[5].smg[2, 3];
       "OUTPUT"."5号梯LEDk" := "IO".elev[5].smg[2, 4];
       "OUTPUT"."5号梯LEDl" := "IO".elev[5].smg[2, 5];
       "OUTPUT"."5号梯LEDm" := "IO".elev[5].smg[2, 6];
       "OUTPUT"."5号梯LEDn" := "IO".elev[5].smg[2, 7];

       "OUTPUT"."5号梯风扇指示" := "IO".elev[5].display.fan;
       "OUTPUT"."5号梯故障指示" := "IO".elev[5].display.error;
       "OUTPUT"."5号梯满载指示" := "IO".elev[5].display.full;
       "OUTPUT"."5号梯照明指示" := "IO".elev[5].display.light;

       "OUTPUT"."5号梯上行指示" := "IO".elev[5].run_disp.up;
       "OUTPUT"."5号梯下行指示" := "IO".elev[5].run_disp.dowm;

       "OUTPUT"."5号梯1级减速制动" := "IO".elev[5].Brake.B1;
       "OUTPUT"."5号梯2级减速制动" := "IO".elev[5].Brake.B2;
       "OUTPUT"."5号梯3级减速制动" := "IO".elev[5].Brake.B3;

       "OUTPUT"."5号梯高速接触器" := "IO".elev[5].ele_speed.H;
       "OUTPUT"."5号梯低速接触器" := "IO".elev[5].ele_speed.L;

       "OUTPUT"."5号梯电机启动信号" := "IO".elev[5].run_enable;
       "OUTPUT"."5号梯上行接触器" := "IO".elev[5].run_contactor.up;
       "OUTPUT"."5号梯下行接触器" := "IO".elev[5].run_contactor.dowm;

       "OUTPUT"."5号梯开门继电器" := "IO".elev[5].door_jdq.open;
       "OUTPUT"."5号梯关门继电器" := "IO".elev[5].door_jdq.close;
   END_REGION
   REGION 6号梯OUTPUT
       "OUTPUT"."6号梯1层按钮指示灯" := "IO".elev[6].ele_in_button[1].light;
       "OUTPUT"."6号梯2层按钮指示灯" := "IO".elev[6].ele_in_button[2].light;
       "OUTPUT"."6号梯3层按钮指示灯" := "IO".elev[6].ele_in_button[3].light;
       "OUTPUT"."6号梯4层按钮指示灯" := "IO".elev[6].ele_in_button[4].light;
       "OUTPUT"."6号梯5层按钮指示灯" := "IO".elev[6].ele_in_button[5].light;
       "OUTPUT"."6号梯6层按钮指示灯" := "IO".elev[6].ele_in_button[6].light;
       "OUTPUT"."6号梯7层按钮指示灯" := "IO".elev[6].ele_in_button[7].light;
       "OUTPUT"."6号梯8层按钮指示灯" := "IO".elev[6].ele_in_button[8].light;
       "OUTPUT"."6号梯9层按钮指示灯" := "IO".elev[6].ele_in_button[9].light;
       "OUTPUT"."6号梯10层按钮指示灯" := "IO".elev[6].ele_in_button[10].light;

       "OUTPUT"."6号梯1层上行呼梯按钮指示灯" := "IO".elev[6].button_out[1, 1].light;
       "OUTPUT"."6号梯2层上行呼梯按钮指示灯" := "IO".elev[6].button_out[1, 2].light;
       "OUTPUT"."6号梯3层上行呼梯按钮指示灯" := "IO".elev[6].button_out[1, 3].light;
       "OUTPUT"."6号梯4层上行呼梯按钮指示灯" := "IO".elev[6].button_out[1, 4].light;
       "OUTPUT"."6号梯5层上行呼梯按钮指示灯" := "IO".elev[6].button_out[1, 5].light;
       "OUTPUT"."6号梯6层上行呼梯按钮指示灯" := "IO".elev[6].button_out[1, 6].light;
       "OUTPUT"."6号梯7层上行呼梯按钮指示灯" := "IO".elev[6].button_out[1, 7].light;
       "OUTPUT"."6号梯8层上行呼梯按钮指示灯" := "IO".elev[6].button_out[1, 8].light;
       "OUTPUT"."6号梯9层上行呼梯按钮指示灯" := "IO".elev[6].button_out[1, 9].light;

       "OUTPUT"."6号梯2层下行呼梯按钮指示灯" := "IO".elev[6].button_out[2, 2].light;
       "OUTPUT"."6号梯3层下行呼梯按钮指示灯" := "IO".elev[6].button_out[2, 3].light;
       "OUTPUT"."6号梯4层下行呼梯按钮指示灯" := "IO".elev[6].button_out[2, 4].light;
       "OUTPUT"."6号梯5层下行呼梯按钮指示灯" := "IO".elev[6].button_out[2, 5].light;
       "OUTPUT"."6号梯6层下行呼梯按钮指示灯" := "IO".elev[6].button_out[2, 6].light;
       "OUTPUT"."6号梯7层下行呼梯按钮指示灯" := "IO".elev[6].button_out[2, 7].light;
       "OUTPUT"."6号梯8层下行呼梯按钮指示灯" := "IO".elev[6].button_out[2, 8].light;
       "OUTPUT"."6号梯9层下行呼梯按钮指示灯" := "IO".elev[6].button_out[2, 9].light;
       "OUTPUT"."6号梯10层下行呼梯按钮指示灯" := "IO".elev[6].button_out[2, 10].light;

       "OUTPUT"."6号梯LEDa" := "IO".elev[6].smg[1, 1];
       "OUTPUT"."6号梯LEDb" := "IO".elev[6].smg[1, 2];
       "OUTPUT"."6号梯LEDc" := "IO".elev[6].smg[1, 3];
       "OUTPUT"."6号梯LEDd" := "IO".elev[6].smg[1, 4];
       "OUTPUT"."6号梯LEDe" := "IO".elev[6].smg[1, 5];
       "OUTPUT"."6号梯LEDf" := "IO".elev[6].smg[1, 6];
       "OUTPUT"."6号梯LEDg" := "IO".elev[6].smg[1, 7];
       "OUTPUT"."6号梯LEDh" := "IO".elev[6].smg[2, 1];
       "OUTPUT"."6号梯LEDi" := "IO".elev[6].smg[2, 2];
       "OUTPUT"."6号梯LEDj" := "IO".elev[6].smg[2, 3];
       "OUTPUT"."6号梯LEDk" := "IO".elev[6].smg[2, 4];
       "OUTPUT"."6号梯LEDl" := "IO".elev[6].smg[2, 5];
       "OUTPUT"."6号梯LEDm" := "IO".elev[6].smg[2, 6];
       "OUTPUT"."6号梯LEDn" := "IO".elev[6].smg[2, 7];

       "OUTPUT"."6号梯风扇指示" := "IO".elev[6].display.fan;
       "OUTPUT"."6号梯故障指示" := "IO".elev[6].display.error;
       "OUTPUT"."6号梯满载指示" := "IO".elev[6].display.full;
       "OUTPUT"."6号梯照明指示" := "IO".elev[6].display.light;

       "OUTPUT"."6号梯上行指示" := "IO".elev[6].run_disp.up;
       "OUTPUT"."6号梯下行指示" := "IO".elev[6].run_disp.dowm;

       "OUTPUT"."6号梯1级减速制动" := "IO".elev[6].Brake.B1;
       "OUTPUT"."6号梯2级减速制动" := "IO".elev[6].Brake.B2;
       "OUTPUT"."6号梯3级减速制动" := "IO".elev[6].Brake.B3;

       "OUTPUT"."6号梯高速接触器" := "IO".elev[6].ele_speed.H;
       "OUTPUT"."6号梯低速接触器" := "IO".elev[6].ele_speed.L;

       "OUTPUT"."6号梯电机启动信号" := "IO".elev[6].run_enable;
       "OUTPUT"."6号梯上行接触器" := "IO".elev[6].run_contactor.up;
       "OUTPUT"."6号梯下行接触器" := "IO".elev[6].run_contactor.dowm;

       "OUTPUT"."6号梯开门继电器" := "IO".elev[6].door_jdq.open;
       "OUTPUT"."6号梯关门继电器" := "IO".elev[6].door_jdq.close;
   END_REGION
END_FUNCTION

FUNCTION "init_up" : Void   // FC2, SCL
{ S7_Optimized_Access := 'TRUE' }
VERSION : 0.1
   VAR_TEMP
      i : Int;
   END_VAR
BEGIN
   FOR #i := 1 TO "ELE_SUM" DO                        
       IF "v_bianliang".dianti[#i].init.kaishi = 1 THEN
           "v_bianliang".dianti[#i].状态指示灯 := 0;
       END_IF;

           CASE "v_bianliang".dianti[#i].init.Init_state OF
               0:
                   REGION 静止态  
                       "v_bianliang".dianti[#i].init.jieshu := 0;
                       "v_bianliang".dianti[#i].init.Init_now_f := 0;
                       "v_bianliang".dianti[#i].Count[2].CV := 0;
                       "v_bianliang".dianti[#i].Count[1].CV := 0;


                           IF NOT "IO".elev[#i].door_inplace.close THEN  
                               "IO".elev[#i].door_jdq.close := 1;
                           ELSE
                               "IO".elev[#i].door_jdq.close := 0;
                           END_IF;

                       IF "v_bianliang".dianti[#i].init.kaishi AND "IO".elev[#i].door_inplace.close THEN
                           IF "v_bianliang".dianti[#i].init.init_fangxiang = 0 THEN 
                               "v_bianliang".dianti[#i].init.Init_state := 1;
                           ELSIF "v_bianliang".dianti[#i].init.init_fangxiang = 1 THEN 
                               "v_bianliang".dianti[#i].init.Init_state := 2;
                           END_IF;
                       END_IF;

                   END_REGION
               1:
                   REGION 初始化方向向下:低速
                       IF #i <> 1 THEN
                           "run_state"(eet_num := #i,
                                       state := "DOWN_L");
                       ELSIF #i = 1 THEN
                           "v_bianliang".dianti[#i].shijian[13].TON(IN := #i = 1,
                                                                    PT := T#0.5S);
                       END_IF;
                       IF "v_bianliang".dianti[#i].shijian[13].Q THEN
                           "run_state"(eet_num := #i,
                                       state := "DOWN_L");
                       END_IF;
                       "IO".elev[#i].run_disp.dowm := 1; 
                       "IO".elev[#i].run_disp.up := 0;
                       IF "IO".elev[#i].bt_limit.bottom1 THEN 
                           "v_bianliang".dianti[#i].init.Init_state := 3;
                       END_IF;
                   END_REGION
               2:
                   REGION 初始化方向向上:低速
                       "run_state"(eet_num := #i,
                                   state := "UP_L");

                       "IO".elev[#i].run_disp.dowm := 0; 
                       "IO".elev[#i].run_disp.up := 1;
                       IF "IO".elev[#i].bt_limit.top1 THEN
                           "v_bianliang".dianti[#i].init.Init_state := 4;
                       END_IF;
                   END_REGION
               3:
                   REGION 折返向上:低速
                       IF "v_bianliang".dianti[#i].gaibian.speed = 1 THEN 

                           "v_bianliang".dianti[#i].shijian[7].TON(IN := "IO".elev[#i].ele_speed.L,
                                                                   PT := T#200MS);
                           IF "v_bianliang".dianti[#i].shijian[7].Q THEN
                               "run_state"(eet_num := #i,
                                           state := "UP_H");
                           END_IF;
                       ELSE
                           "run_state"(eet_num := #i,
                                       state := "UP_L");
                       END_IF;

                       "IO".elev[#i].run_disp.dowm := 0;
                       "IO".elev[#i].run_disp.up := 1;

                       "v_bianliang".dianti[#i].Count[1].CTU(CU := "IO".elev[#i].run_contactor.up AND "IO".elev[#i].direction.up AND "IO".elev[#i].direction.down,
                                                             PV := "FlOOR_TOP",
                                                             CV => "v_bianliang".dianti[#i].init.Init_now_f);

                       IF "v_bianliang".dianti[#i].init.Init_now_f = "v_bianliang".dianti[#i].init.mubiao_floor THEN 
                           "v_bianliang".dianti[#i].init.Init_state := 5;
                       END_IF;
                   END_REGION ;
               4:
                   REGION 折返向下:低速
                       IF "v_bianliang".dianti[#i].gaibian.speed = 1 THEN 

                           "v_bianliang".dianti[#i].shijian[7].TON(IN := "IO".elev[#i].ele_speed.L,
                                                                   PT := T#200MS);
                           IF "v_bianliang".dianti[#i].shijian[7].Q THEN
                               "run_state"(eet_num := #i,
                                           state := "DOWN_H");
                           END_IF;
                       ELSE
                           "run_state"(eet_num := #i,
                                       state := "DOWN_L");
                       END_IF;

                       "IO".elev[#i].run_disp.dowm := 1;
                       "IO".elev[#i].run_disp.up := 0;

                       "v_bianliang".dianti[#i].Count[2].CTU(CU := "IO".elev[#i].run_contactor.dowm AND "IO".elev[#i].direction.up AND "IO".elev[#i].direction.down,
                                                             PV := "FlOOR_TOP",
                                                             CV => "v_bianliang".dianti[#i].init.Init_now_f);

                       IF ("FlOOR_TOP" + 1 - "v_bianliang".dianti[#i].init.Init_now_f) = "v_bianliang"."dianti"[#i].init.mubiao_floor THEN
                           "v_bianliang".dianti[#i].init.Init_state := 5;
                       END_IF;
                   END_REGION
               5:
                   REGION 静止态
                       "run_state"(eet_num := #i,
                                   state := "STATIC");

                       "IO".elev[#i].run_disp.dowm := 0; 
                       "IO".elev[#i].run_disp.up := 0;

                       "v_bianliang".dianti[#i].Floor_handle.dangqian_floor := "v_bianliang".dianti[#i].init.mubiao_floor;//将初始化到达楼层赋值给全局的楼层计数
                       "v_bianliang".dianti[#i].Count[3].CV := "v_bianliang".dianti[#i].init.mubiao_floor;

                       "v_bianliang".dianti[#i].init.kaishi := 0;
                       "v_bianliang".dianti[#i].init.jieshu := 1;

                       "v_bianliang".dianti[#i].init.Init_state := 0;

                       RESET_TIMER("v_bianliang".dianti[#i].shijian[7]); 
                       RESET_TIMER("v_bianliang".dianti[#i].shijian[13]);
                   END_REGION
           END_CASE;
   END_FOR;

   FOR #i := 1 TO "ELE_SUM" DO
       IF "v_bianliang".dianti[#i].init.jieshu THEN //若电梯初始化完毕，则计数标志cnt+1
           "v_bianliang".cnt_wancheng += 1;
       END_IF;
   END_FOR;
   FOR #i := "ELE_SUM" TO 1 BY -1 DO
       IF "v_bianliang".dianti[#i].cuowu.REP_deal AND NOT "v_bianliang".dianti[#i].cuowu.tag_REPR THEN //若有电梯检修，则计数标志cnt+1
           "v_bianliang".cnt_wancheng += 1;
       END_IF;
       "v_bianliang".dianti[#i].cuowu.tag_REPR := "v_bianliang".dianti[#i].cuowu.REP_deal;
   END_FOR;
   IF "v_bianliang".cnt_wancheng = "ELE_SUM" THEN 
       "IO".plc_ready := 1;
   END_IF;
   FOR #i := 1 TO "ELE_SUM" DO
       IF "v_bianliang".dianti[#i].init.jieshu THEN 
           "v_bianliang".dianti[#i].yunxing_chuli.yunxu_run := 1;
       END_IF;
   END_FOR;
END_FUNCTION

FUNCTION "init_signal" : Void   // FC3, SCL
{ S7_Optimized_Access := 'TRUE' }
VERSION : 0.1
   VAR_TEMP
      i : Int;
      j : Int;
      res_cnt : Int;
   END_VAR
BEGIN
   "Res"(CLK := "IO".software_autorun OR "v_bianliang".autorun OR "v_bianliang".初始信号 );

   IF "Res".Q THEN                                       
       "v_bianliang".zidongyuxing_cnt := "v_bianliang".zidongyuxing_cnt  + 1;
       FOR #i := 1 TO "ELE_SUM" DO
           "v_bianliang".dianti[#i].init.init_fangxiang := "v_bianliang".dianti[#i].gaibian.init_dir;
           "v_bianliang".dianti[#i].init.mubiao_floor := "v_bianliang".dianti[#i].gaibian.init_aimf;
           "run_state"(eet_num := #i,
                           state := "STATIC");
           "v_bianliang".dianti[#i].init.Init_state := 0;
       END_FOR;
   END_IF;

   IF "Res".Q AND "v_bianliang".zidongyuxing_cnt  = 1 THEN                 //第一次初始化

       FOR #i := 1 TO "ELE_SUM" DO
           "v_bianliang".dianti[#i].init.kaishi := 1;
       END_FOR;

   END_IF;
   //1
   IF "Res".Q AND "v_bianliang".zidongyuxing_cnt  = 2 THEN             //第二次初始化
       "IO".plc_ready := 0;                         

       "init"();//进行相关中间变量复位

       "v_bianliang".mode_choice += 1; 
       FOR #i := 1 TO "ELE_SUM" DO
           "v_bianliang".dianti[#i].init.kaishi := 1;        //再次发出初始化信号
       END_FOR;
   END_IF;
   //2
   IF "Res".Q AND "v_bianliang".zidongyuxing_cnt = 3 THEN             //第三次初始化
       "IO".plc_ready := 0;                         

       "init"();//进行相关中间变量复位

       "v_bianliang".mode_choice += 1;
       FOR #i := 1 TO "ELE_SUM" DO
           "v_bianliang".dianti[#i].init.kaishi := 1;        
       END_FOR;
   END_IF;
   //3
   IF "Res".Q AND "v_bianliang".zidongyuxing_cnt = 4 THEN             //第四次初始化
       "IO".plc_ready := 0;

       "init"(); 

       "v_bianliang".mode_choice += 1;
       FOR #i := 1 TO "ELE_SUM" DO
           "v_bianliang".dianti[#i].init.kaishi := 1;        
       END_FOR;
   END_IF;
END_FUNCTION

FUNCTION "show_F" : Void   // FC4, SCL
{ S7_Optimized_Access := 'TRUE' }
VERSION : 0.1
   VAR_TEMP
      i : Int;
   END_VAR
BEGIN
   FOR #i := 1 TO "ELE_SUM" DO
       IF "v_bianliang".dianti[#i].yunxing_chuli.yunxu_run THEN

           IF "IO".elev[#i].run_contactor.up AND NOT "v_bianliang".dianti[#i].Floor_handle.tag_1 THEN
               "v_bianliang".dianti[#i].Count[3].CV := "v_bianliang".dianti[#i].Count[3].CV - 1;
           END_IF;
           "v_bianliang".dianti[#i].Floor_handle.tag_1 := "IO".elev[#i].run_contactor.up;


           IF "IO".elev[#i].run_contactor.dowm AND NOT "v_bianliang".dianti[#i].Floor_handle.tag_2 THEN
               "v_bianliang".dianti[#i].Count[3].CV := "v_bianliang".dianti[#i].Count[3].CV + 1;
           END_IF;
           "v_bianliang".dianti[#i].Floor_handle.tag_2 := "IO".elev[#i].run_contactor.dowm;


           "v_bianliang".dianti[#i].Count[3].CTUD(CU := "IO".elev[#i].run_contactor.up AND "IO".elev[#i].direction.up,
                                      CD := "IO".elev[#i].run_contactor.dowm AND "IO".elev[#i].direction.down,
                                      PV := "FlOOR_TOP",
                                      CV => "v_bianliang".dianti[#i].Floor_handle.dangqian_floor);


           "smg_display"(Number := "v_bianliang".dianti[#i].Floor_handle.dangqian_floor MOD 10, 
                 Output_A => "IO".elev[#i].smg[1, 1],
                 Output_B => "IO".elev[#i].smg[1, 2],
                 Output_C => "IO".elev[#i].smg[1, 3],
                 Output_D => "IO".elev[#i].smg[1, 4],
                 Output_E => "IO".elev[#i].smg[1, 5],
                 Output_F => "IO".elev[#i].smg[1, 6],
                 Output_G => "IO".elev[#i].smg[1, 7]);

           "smg_display"(Number := "v_bianliang".dianti[#i].Floor_handle.dangqian_floor / 10, 
                 Output_A => "IO".elev[#i].smg[2, 1],
                 Output_B => "IO".elev[#i].smg[2, 2],
                 Output_C => "IO".elev[#i].smg[2, 3],
                 Output_D => "IO".elev[#i].smg[2, 4],
                 Output_E => "IO".elev[#i].smg[2, 5],
                 Output_F => "IO".elev[#i].smg[2, 6],
                 Output_G => "IO".elev[#i].smg[2, 7]);
       END_IF;
   END_FOR;
END_FUNCTION

FUNCTION "smg_display" : Void   // FC5, SCL
{ S7_Optimized_Access := 'TRUE' }
VERSION : 0.1
   VAR_INPUT
      Number : Int;
   END_VAR
   VAR_OUTPUT
      Output_A : Bool;
      Output_B : Bool;
      Output_C : Bool;
      Output_D : Bool;
      Output_E : Bool;
      Output_F : Bool;
      Output_G : Bool;
   END_VAR
BEGIN
   CASE #Number OF
       0:
           #Output_A := 1;
           #Output_B := 1;
           #Output_C := 1;
           #Output_D := 1;
           #Output_E := 1;
           #Output_F := 1;
           #Output_G := 0;
       1:
           #Output_A := 0;
           #Output_B := 1;
           #Output_C := 1;
           #Output_D := 0;
           #Output_E := 0;
           #Output_F := 0;
           #Output_G := 0;
       2:
           #Output_A := 1;
           #Output_B := 1;
           #Output_C := 0;
           #Output_D := 1;
           #Output_E := 1;
           #Output_F := 0;
           #Output_G := 1;
       3:
           #Output_A := 1;
           #Output_B := 1;
           #Output_C := 1;
           #Output_D := 1;
           #Output_E := 0;
           #Output_F := 0;
           #Output_G := 1;
       4:
           #Output_A := 0;
           #Output_B := 1;
           #Output_C := 1;
           #Output_D := 0;
           #Output_E := 0;
           #Output_F := 1;
           #Output_G := 1;
       5:
           #Output_A := 1;
           #Output_B := 0;
           #Output_C := 1;
           #Output_D := 1;
           #Output_E := 0;
           #Output_F := 1;
           #Output_G := 1;
       6:
           #Output_A := 1;
           #Output_B := 0;
           #Output_C := 1;
           #Output_D := 1;
           #Output_E := 1;
           #Output_F := 1;
           #Output_G := 1;
       7:
           #Output_A := 1;
           #Output_B := 1;
           #Output_C := 1;
           #Output_D := 0;
           #Output_E := 0;
           #Output_F := 0;
           #Output_G := 0;
       8:
           #Output_A := 1;
           #Output_B := 1;
           #Output_C := 1;
           #Output_D := 1;
           #Output_E := 1;
           #Output_F := 1;
           #Output_G := 1;
       9:
           #Output_A := 1;
           #Output_B := 1;
           #Output_C := 1;
           #Output_D := 1;
           #Output_E := 0;
           #Output_F := 1;
           #Output_G := 1;
   END_CASE;
END_FUNCTION

FUNCTION "CALL_ELE" : Void   // FC6, SCL
{ S7_Optimized_Access := 'TRUE' }
VERSION : 0.1
   VAR_TEMP
      i : Int;
      j : Int;
   END_VAR
BEGIN
   REGION 内呼处理
       FOR #i := 1 TO "ELE_SUM" DO

           FOR #j := 1 TO "FlOOR_TOP" DO

               "nei_hu"(i:=#i,
                        j:=#j);

           END_FOR;

       END_FOR;
   END_REGION 

   REGION 外呼录入    
       FOR #i := 1 TO "ELE_SUM" DO
           FOR #j := 1 TO "FlOOR_TOP" - 1 DO//上呼录入
               IF "IO".elev[#i].button_out[1, #j].state AND NOT "IO".elev[#i].button_out[1, #j].p THEN
                   "v_bianliang".anniu_waibu[1, #j] := 1;
                   "IO".elev[#i].button_out[1, #j].light := 1;
                   IF "v_bianliang".dianti[#i].Floor_handle.dangqian_floor <> #j THEN
                       "v_bianliang".over_tim[1, #j] := "v_bianliang".all_time.min * 60 + "v_bianliang".all_time.sec;//结束时间
                   END_IF;
               END_IF;
               "IO".elev[#i].button_out[1, #j].p := "IO".elev[#i].button_out[1, #j].state;
               IF "v_bianliang".anniu_waibu[1, #j] = 0 THEN
                   "IO".elev[#i].button_out[1, #j].light := 0;
               END_IF;
           END_FOR;

           FOR #j := 2 TO "FlOOR_TOP" DO//下呼录入
                   IF "IO".elev[#i].button_out[2, #j].state AND NOT "IO".elev[#i].button_out[2, #j].p THEN
                       "v_bianliang".anniu_waibu[2, #j] := 1;
                       "IO".elev[#i].button_out[2, #j].light := 1;
                       IF "v_bianliang".dianti[#i].Floor_handle.dangqian_floor <> #j THEN
                           "v_bianliang".over_tim[2, #j] := "v_bianliang".all_time.min * 60 + "v_bianliang".all_time.sec;//结束时间
                       END_IF;
                   END_IF;
                   "IO".elev[#i].button_out[2, #j].p := "IO".elev[#i].button_out[2, #j].state;
                   IF "v_bianliang".anniu_waibu[2, #j] = 0 THEN
                       "IO".elev[#i].button_out[2, #j].light := 0;
                   END_IF;
           END_FOR;
       END_FOR;
   END_REGION

   // REGION 单体外呼录入    
   //     FOR #i := 1 TO "ELE_SUM" DO//使用这个要把群控屏蔽
   //         FOR #j := 1 TO "FlOOR_TOP" - 1 DO//上呼录入
   //             IF "IO".elev[#i].button_out[1, #j].state AND NOT "IO".elev[#i].button_out[1, #j].p THEN
   //                 "v_bianliang"."dianti"[#i].anniu_luru.waibu_anniu[1, #j] := 1;
   //                 "IO".elev[#i].button_out[1, #j].light := 1;
   //             END_IF;
   //             "IO".elev[#i].button_out[1, #j].p := "IO".elev[#i].button_out[1, #j].state;
   //             IF "v_bianliang"."dianti"[#i].anniu_luru.waibu_anniu[1, #j] = 0 THEN
   //                 "IO".elev[#i].button_out[1, #j].light := 0;
   //             END_IF;
   //         END_FOR;

   //         FOR #j := 2 TO "FlOOR_TOP" DO//下呼录入
   //             IF "IO".elev[#i].button_out[2, #j].state AND NOT "IO".elev[#i].button_out[2, #j].p THEN
   //                 "v_bianliang"."dianti"[#i].anniu_luru.waibu_anniu[2, #j] := 1;
   //                 "IO".elev[#i].button_out[2, #j].light := 1;
   //             END_IF;
   //             "IO".elev[#i].button_out[2, #j].p := "IO".elev[#i].button_out[2, #j].state;
   //             IF "v_bianliang"."dianti"[#i].anniu_luru.waibu_anniu[2, #j] = 0 THEN
   //                 "IO".elev[#i].button_out[2, #j].light := 0;
   //             END_IF;
   //         END_FOR;
   //     END_FOR;
   // END_REGION

   // REGION 开关门录入
   //     FOR #i := 1 TO "ELE_SUM" DO//电梯开门
   //         IF ("IO".elev[#i].door_open.state AND NOT "IO".elev[#i].door_open.p) OR (NOT "IO".elev[#i].door_open.state AND "IO".elev[#i].door_open.p) THEN
   //             "v_bianliang".dianti[#i].yunxing_chuli.run_state := 7;
   //         END_IF;
   //             "IO".elev[#i].door_open.p := "IO".elev[#i].door_open.state;
   //     END_FOR;
   //     // FOR #i := 1 TO "ELE_SUM" DO//电梯关门
   //     //     IF ("IO".elev[#i].btn_close.state AND NOT "IO".elev[#i].btn_close.p) OR (NOT "IO".elev[#i].btn_close.state AND "IO".elev[#i].btn_close.p) THEN
   //     //         "v_bianliang".dianti[#i].yunxing_chuli.run_state := 8;
   //     //     END_IF;
   //     //     "IO".elev[#i].btn_close.p := "IO".elev[#i].btn_close.state;
   //     // END_FOR;
   // END_REGION
END_FUNCTION

FUNCTION "timer" : Void   // FC7, SCL
{ S7_Optimized_Access := 'TRUE' }
VERSION : 0.1
   VAR_TEMP
      i : Int;
   END_VAR
BEGIN
   // IF "variable".interrupt.f_1ms = 1 THEN
   //     "variable".interrupt.f_1ms := 0;
   //     "variable".interrupt.cnt_100ms += 1;
   //     IF "variable".interrupt.cnt_100ms = 100 THEN
   //         "variable".interrupt.cnt_100ms := 0;
   //         "variable".interrupt.f_100ms := 1;
   //     END_IF;
   // END_IF;

   FOR #i := 1 TO "ELE_SUM" DO
       IF "v_bianliang".dianti[#i].interrupt.f_1ms = 1 THEN
           "v_bianliang".dianti[#i].interrupt.f_1ms := 0;
           "v_bianliang".dianti[#i].interrupt.cnt_100ms += 1;
           IF "v_bianliang".dianti[#i].interrupt.cnt_100ms = 100 THEN
               "v_bianliang".dianti[#i].interrupt.cnt_100ms := 0;
               "v_bianliang".dianti[#i].interrupt.f_100ms := 1;
           END_IF;
       END_IF;
   END_FOR;
END_FUNCTION

FUNCTION "init" : Void   // FC8, SCL
{ S7_Optimized_Access := 'TRUE' }
VERSION : 0.1
   VAR_TEMP
      i : Int;
      j : Int;
   END_VAR
BEGIN
       REGION 进行相关中间变量复位    
           "v_bianliang".cnt_wancheng := 0;//完成初始化的电梯计数置0
           "v_bianliang".zuiyou_dianti := 0;
           FOR #i := 1 TO "ELE_SUM" DO
               "v_bianliang".dianti[#i].cuowu.tag_REPR := 0;
               "v_bianliang".dianti[#i].yunxing_chuli.yunxu_run := 0; //电梯禁止运行
               "v_bianliang".dianti[#i].yunxing_chuli.run_state := 0; //运行状态机为静止态
               "v_bianliang".dianti[#i].yunxing_chuli.uopdown_state := 0; //上下行状态为静止
               FOR #j := 1 TO "FlOOR_TOP" DO //外呼虚拟楼层和内呼信号置0
                   "v_bianliang".dianti[#i].anniu_luru.neibu_anniu[#j] := 0;
                   "v_bianliang".dianti[#i].anniu_luru.waibu_anniu[1, #j] := 0;
                   "v_bianliang".dianti[#i].anniu_luru.waibu_anniu[2, #j] := 0;
               END_FOR;
               "v_bianliang".dianti[#i].Weight_handle.shiji_load := 0;//载重相关变量清0
               "v_bianliang".dianti[#i].Weight_handle.jiangyao_chaozhong := 0;
               "v_bianliang".time_min[#i] := 0;//群控相关变量清0
               "v_bianliang".dianti[#i].qunkong.TH := 0;
               RESET_TIMER("v_bianliang".dianti[#i].shijian[1]);
               RESET_TIMER("v_bianliang".dianti[#i].shijian[2]);
               RESET_TIMER("v_bianliang".dianti[#i].shijian[3]);
               RESET_TIMER("v_bianliang".dianti[#i].shijian[4]);
               RESET_TIMER("v_bianliang".dianti[#i].shijian[5]);
               RESET_TIMER("v_bianliang".dianti[#i].shijian[6]);
               RESET_TIMER("v_bianliang".dianti[#i].shijian[7]);
               RESET_TIMER("v_bianliang".dianti[#i].shijian[8]);
               RESET_TIMER("v_bianliang".dianti[#i].shijian[9]);
               RESET_TIMER("v_bianliang".dianti[#i].shijian[10]);
               RESET_TIMER("v_bianliang".dianti[#i].shijian[11]);
               RESET_TIMER("v_bianliang".dianti[#i].shijian[12]);
           END_FOR;
           FOR #i := 1 TO "FlOOR_TOP" DO
               "v_bianliang".anniu_waibu[1, #i] := 0;
               "v_bianliang".anniu_waibu[2, #i] := 0;
           END_FOR;
       END_REGION

       REGION 进行PLC输出信号复位 


           REGION 其余信号
               FOR #i := 1 TO "ELE_SUM" DO
                   "IO".elev[#i].ele_in_button[1].light := 0;
                   "IO".elev[#i].ele_in_button[2].light := 0;
                   "IO".elev[#i].ele_in_button[3].light := 0;
                   "IO".elev[#i].ele_in_button[4].light := 0;
                   "IO".elev[#i].ele_in_button[5].light := 0;
                   "IO".elev[#i].ele_in_button[6].light := 0;
                   "IO".elev[#i].ele_in_button[7].light := 0;
                   "IO".elev[#i].ele_in_button[8].light := 0;
                   "IO".elev[#i].ele_in_button[9].light := 0;
                   "IO".elev[#i].ele_in_button[10].light := 0;

                   "IO".elev[#i].button_out[1, 1].light := 0;
                   "IO".elev[#i].button_out[1, 2].light := 0;
                   "IO".elev[#i].button_out[1, 3].light := 0;
                   "IO".elev[#i].button_out[1, 4].light := 0;
                   "IO".elev[#i].button_out[1, 5].light := 0;
                   "IO".elev[#i].button_out[1, 6].light := 0;
                   "IO".elev[#i].button_out[1, 7].light := 0;
                   "IO".elev[#i].button_out[1, 8].light := 0;
                   "IO".elev[#i].button_out[1, 9].light := 0;

                   "IO".elev[#i].button_out[2, 2].light := 0;
                   "IO".elev[#i].button_out[2, 3].light := 0;
                   "IO".elev[#i].button_out[2, 4].light := 0;
                   "IO".elev[#i].button_out[2, 5].light := 0;
                   "IO".elev[#i].button_out[2, 6].light := 0;
                   "IO".elev[#i].button_out[2, 7].light := 0;
                   "IO".elev[#i].button_out[2, 8].light := 0;
                   "IO".elev[#i].button_out[2, 9].light := 0;
                   "IO".elev[#i].button_out[2, 10].light := 0;

                   "IO".elev[#i].smg[1, 1] := 0;
                   "IO".elev[#i].smg[1, 2] := 0;
                   "IO".elev[#i].smg[1, 3] := 0;
                   "IO".elev[#i].smg[1, 4] := 0;
                   "IO".elev[#i].smg[1, 5] := 0;
                   "IO".elev[#i].smg[1, 6] := 0;
                   "IO".elev[#i].smg[1, 7] := 0;
                   "IO".elev[#i].smg[2, 1] := 0;
                   "IO".elev[#i].smg[2, 2] := 0;
                   "IO".elev[#i].smg[2, 3] := 0;
                   "IO".elev[#i].smg[2, 4] := 0;
                   "IO".elev[#i].smg[2, 5] := 0;
                   "IO".elev[#i].smg[2, 6] := 0;
                   "IO".elev[#i].smg[2, 7] := 0;

                   "IO".elev[#i].display.fan := 0;
                   "IO".elev[#i].display.error := 0;
                   "IO".elev[#i].display.full := 0;
                   "IO".elev[#i].display.light := 0;

                   "IO".elev[#i].run_disp.up := 0;
                   "IO".elev[#i].run_disp.dowm := 0;

                   "IO".elev[#i].Brake.B1 := 0;
                   "IO".elev[#i].Brake.B2 := 0;
                   "IO".elev[#i].Brake.B3 := 0;

                   "IO".elev[#i].ele_speed.H := 0;
                   "IO".elev[#i].ele_speed.L := 0;

                   "IO".elev[#i].run_enable := 0;
                   "IO".elev[#i].run_contactor.up := 0;
                   "IO".elev[#i].run_contactor.dowm := 0;

                   "IO".elev[#i].door_jdq.open := 0;
                   "IO".elev[#i].door_jdq.close := 0;


               END_FOR;
           END_REGION

       END_REGION
END_FUNCTION

FUNCTION "run_state" : Void   // FC9, SCL
{ S7_Optimized_Access := 'TRUE' }
VERSION : 0.1
   VAR_INPUT
      eet_num : Int;
      state : Int;
   END_VAR
BEGIN
   CASE #state OF
       0: REGION 静止
               "IO".elev[#eet_num].ele_speed.H := 0;
               "IO".elev[#eet_num].ele_speed.L := 0;
               "IO".elev[#eet_num].run_enable := 0;
               "IO".elev[#eet_num].run_contactor.up := 0;
               "IO".elev[#eet_num].run_contactor.dowm := 0;
               "IO".elev[#eet_num].door_jdq.open := 0;
               "IO".elev[#eet_num].door_jdq.close := 0;
           END_REGION 
       1: REGION 上行高速
               "IO".elev[#eet_num].ele_speed.H := 1;
               "IO".elev[#eet_num].ele_speed.L := 0;
               "IO".elev[#eet_num].run_enable := 1;
               "IO".elev[#eet_num].run_contactor.up := 1;
               "IO".elev[#eet_num].run_contactor.dowm := 0;
               "IO".elev[#eet_num].door_jdq.open := 0;
               "IO".elev[#eet_num].door_jdq.close := 0;
           END_REGION
       2: REGION 上行低速
               "IO".elev[#eet_num].ele_speed.H := 0;
               "IO".elev[#eet_num].ele_speed.L := 1;
               "IO".elev[#eet_num].run_enable := 1;
               "IO".elev[#eet_num].run_contactor.up := 1;
               "IO".elev[#eet_num].run_contactor.dowm := 0;
               "IO".elev[#eet_num].door_jdq.open := 0;
               "IO".elev[#eet_num].door_jdq.close := 0;
           END_REGION
       3: REGION 下行高速
               "IO".elev[#eet_num].ele_speed.H := 1;
               "IO".elev[#eet_num].ele_speed.L := 0;
               "IO".elev[#eet_num].run_enable := 1;
               "IO".elev[#eet_num].run_contactor.up := 0;
               "IO".elev[#eet_num].run_contactor.dowm := 1;
               "IO".elev[#eet_num].door_jdq.open := 0;
               "IO".elev[#eet_num].door_jdq.close := 0;
           END_REGION
       4: REGION 下行低速
               "IO".elev[#eet_num].ele_speed.H := 0;
               "IO".elev[#eet_num].ele_speed.L := 1;
               "IO".elev[#eet_num].run_enable := 1;
               "IO".elev[#eet_num].run_contactor.up := 0;
               "IO".elev[#eet_num].run_contactor.dowm := 1;
               "IO".elev[#eet_num].door_jdq.open := 0;
               "IO".elev[#eet_num].door_jdq.close := 0;
           END_REGION
       5: REGION 开门
               "IO".elev[#eet_num].ele_speed.H := 0;
               "IO".elev[#eet_num].ele_speed.L := 0;
               "IO".elev[#eet_num].run_enable := 0;
               "IO".elev[#eet_num].run_contactor.up := 0;
               "IO".elev[#eet_num].run_contactor.dowm := 0;
               "IO".elev[#eet_num].door_jdq.open := 1;
               "IO".elev[#eet_num].door_jdq.close := 0;
           END_REGION
       6: REGION 关门
               "IO".elev[#eet_num].ele_speed.H := 0;
               "IO".elev[#eet_num].ele_speed.L := 0;
               "IO".elev[#eet_num].run_enable := 0;
               "IO".elev[#eet_num].run_contactor.up := 0;
               "IO".elev[#eet_num].run_contactor.dowm := 0;
               "IO".elev[#eet_num].door_jdq.open := 0;
               "IO".elev[#eet_num].door_jdq.close := 1;
           END_REGION
       7: REGION 高速切低速
               "IO".elev[#eet_num].ele_speed.H := 0;
               "IO".elev[#eet_num].ele_speed.L := 1;
           END_REGION
       8: REGION 低速切高速
               "IO".elev[#eet_num].ele_speed.H := 1;
               "IO".elev[#eet_num].ele_speed.L := 0;
           END_REGION
   END_CASE;
END_FUNCTION

FUNCTION "Indicate" : Void   // FC10, SCL
{ S7_Optimized_Access := 'TRUE' }
VERSION : 0.1
   VAR_TEMP
      i : Int;
   END_VAR
BEGIN
   FOR #i := 1 TO "ELE_SUM" DO
       IF "v_bianliang".dianti[#i].yunxing_chuli.yunxu_run THEN
           REGION 上下行显示
               IF "v_bianliang".dianti[#i].yunxing_chuli.uopdown_state = 0 THEN
                   "IO".elev[#i].run_disp.dowm := 0;
                   "IO".elev[#i].run_disp.up := 0;
               ELSIF "v_bianliang".dianti[#i].yunxing_chuli.uopdown_state = 1 THEN
                   "IO".elev[#i].run_disp.dowm := 0;
                   "IO".elev[#i].run_disp.up := 1;
               ELSIF "v_bianliang".dianti[#i].yunxing_chuli.uopdown_state = 2 THEN
                   "IO".elev[#i].run_disp.dowm := 1;
                   "IO".elev[#i].run_disp.up := 0;
               END_IF;
           END_REGION

           REGION 照明与风扇显示
               IF "v_bianliang".dianti[#i].Weight_handle.shiji_load = 0 THEN 
                   "IO".elev[#i].display.fan := 0;
                   "IO".elev[#i].display.light := 0;
               ELSE
                   "IO".elev[#i].display.fan := 1;
                   "IO".elev[#i].display.light := 1;
               END_IF;
           END_REGION

           REGION 超载显示
               IF "v_bianliang".dianti[#i].Weight_handle.chaozhongxinhao THEN
                   "IO".elev[#i].display.full := 1;
               ELSE
                   "IO".elev[#i].display.full := 0;
               END_IF;
           END_REGION
       END_IF;
   END_FOR;
END_FUNCTION

FUNCTION "signal_check" : Void   // FC11, SCL
{ S7_Optimized_Access := 'TRUE' }
VERSION : 0.1
   VAR_TEMP
      i : Int;
      state : Int;
   END_VAR
BEGIN
   FOR #i := 1 TO "ELE_SUM" DO

